(* IEC 61131-3 sources: daoli-st-library/DL_MathData (part 2) *)

(* ---- FC_DL_DtlStringConv.st ---- *)
(*
  ==================================================================
  组件名 Component  : FC_DL_DtlStringConv
  分类   Category   : DL_MathData
  复杂度 Complexity  : 中
  版本   Version    : 1.0.0
  功能   Purpose    : 日期时间 ↔ ASCII 串双向转换。定长 19 字符格式
                      'YYYY-MM-DD HH:MM:SS'。eStrToComp：串 → 六分量（分隔符
                      与数字位逐一校验，FIND 数字表解码）；eCompToStr：六分量
                      → 串（数字查表装配）。超长按 19 截断评估并置 bTrunc
                      （255 截断标志语义：入串超库上限 255 或超定长均置位）。
                      LGF Converter 组 DTL↔String 语义 clean-room。
  来源   Source     : T2-1-lgf-converter（LGF Converter 组 DTL↔String 语义）
  溯源   Origin     : 定长日期串装配/解析为公开工程语义，clean-room 自研实现，
                      未复制 LGF 或任何厂商私有库源码。
  平台   Platform   : 纯 IEC 61131-3（Standard.library: LEN / MID / CONCAT /
                      FIND，无私有库）
  分工声明 Split     : 与 FC_DL_AsciiFrameParse 分工——后者做 STX/ETX 仪表
                      帧解析，本件做定长日期时间串双向转换。
  作者   Author     : 道莅代码库 · PLC 编程专家（R59）
  ------------------------------------------------------------------
  边界 Boundary     :
                      一 值域闸（eCompToStr）：年 1970..2999 / 月 1..12 /
                         日 1..31 / 时 0..23 / 分秒 0..59，越域置 bError；
                      二 格式闸（eStrToComp）：定长 19、分隔符位置（5/8 =
                         '-'，11 = ' '，14/17 = ':'）、数字位非数字 → bError；
                      三 255 截断标志：LEN > 19 按前 19 位截断评估并置
                         bTrunc（信息级），LEN > 255 直接置 bError；
                      四 无除法无浮点（纯整数与串操作，无除零/非有限风险）；
                      五 无全局变量、无外部变量声明、无物理地址寻址。
  修订记录 Revision  :
    2026-11-21  v1.0.0  R59 首版（批 2 · 序号 6）
  ==================================================================
*)

TYPE E_DL_DtcMode :
(
    eStrToComp := 0, // 串 → 六分量 / the string to components direction
    eCompToStr := 1  // 六分量 → 串 / the components to string direction
);
END_TYPE

FUNCTION FC_DL_DtlStringConv : BOOL
VAR_INPUT
    eMode   : E_DL_DtcMode; // 转换方向枚举 [-] / the conversion direction enum
    sIn     : STRING(255) := ''; // 入串（eStrToComp 方向）[-] / the input string, the to components entry
    nYear   : DINT := 2000; // 年分量 [年]，域 1970..2999，eCompToStr 方向 / the year component
    nMonth  : DINT := 1;    // 月分量 [月]，域 1..12 / the month component
    nDay    : DINT := 1;    // 日分量 [日]，域 1..31 / the day component
    nHour   : DINT := 0;    // 时分量 [时]，域 0..23 / the hour component
    nMinute : DINT := 0;    // 分分量 [分]，域 0..59 / the minute component
    nSecond : DINT := 0;    // 秒分量 [秒]，域 0..59 / the second component
END_VAR
VAR_OUTPUT
    sOut    : STRING(23) := ''; // 出串 'YYYY-MM-DD HH:MM:SS' [-] / the output string, the fixed format
    oYear   : DINT := 0;   // 年分量输出 [年] / the year outlet
    oMonth  : DINT := 0;   // 月分量输出 [月] / the month outlet
    oDay    : DINT := 0;   // 日分量输出 [日] / the day outlet
    oHour   : DINT := 0;   // 时分量输出 [时] / the hour outlet
    oMinute : DINT := 0;   // 分分量输出 [分] / the minute outlet
    oSecond : DINT := 0;   // 秒分量输出 [秒] / the second outlet
    bValid  : BOOL := FALSE; // 结果可用标志 [-] / the result usable flag
    bTrunc  : BOOL := FALSE; // 截断标志（入串超定长 19 按前 19 位评估）[-] / the truncation flag, the long input evaluated by the first nineteen
    bError  : BOOL := FALSE; // 故障标志（格式/值域/超 255）[-] / the fault flag
END_VAR
VAR CONSTANT
    DL_DTC_DIGITS : STRING(10) := '0123456789'; // 数字字符表（FIND 解码基准）/ the digit table for the FIND decoding
    DL_DTC_LENFIX : DINT := 19; // 定长 [字符] / the fixed length
    DL_DTC_LENMAX : DINT := 255; // 库串上限 [字符] / the library string cap
END_VAR
VAR
    nLen   : DINT;  // 入串长度 [字符] / the input length
    sCh    : STRING(1); // 单字符工作量 [-] / the one char work value
    nPos   : DINT;  // 字表命中位（0 = 非数字）[位] / the table hit position, zero means non digit
    nI     : DINT;  // 数字位遍历索引 [位] / the digit position index
    nJ     : DINT;  // 字段遍历索引 [个] / the field index
    nVal   : DINT;  // 字段解析值工作量 [-] / the field parsed value work
    nDiv   : DINT;  // 位除子工作量（10 的幂，DINT 整除取位）[-] / the digit divisor, a power of ten
    aVal   : ARRAY[0..5] OF DINT; // 六分量装配工作数组 / the six component work array
    aField : ARRAY[0..5] OF DINT; // 六字段起始位组（1 基）/ the six field start positions, one based
    aWidth : ARRAY[0..5] OF DINT; // 六字段宽度组 [字符] / the six field widths
    aSep   : ARRAY[0..5] OF STRING(1); // 字段间分隔符组（末项空）/ the separators, the last empty
    bNeg   : BOOL;  // 保留（本件无符号语义，恒假）[-] / reserved, constant false
END_VAR

// 段 1｜返回值与输出预置（四段式第一段，R45）/ segment 1, preset the return and the outputs
FC_DL_DtlStringConv := FALSE; // 受理预置假 / preset the accepted false
sOut := ''; // 出串预置空 / preset the output empty
oYear := 0; oMonth := 0; oDay := 0; // 分量输出预置零 / preset the outlets zero
oHour := 0; oMinute := 0; oSecond := 0; // 分量输出预置零 / preset the outlets zero
bValid := FALSE; // 有效预置假 / preset the valid false
bTrunc := FALSE; // 截断预置假 / preset the trunc false
bError := FALSE; // 故障预置假 / preset the fault false
bNeg := FALSE; // 保留位恒假 / the reserved constant false

// 段 2｜方向一：串 → 六分量（格式闸 + 数字表解码 + 值域闸）/ segment 2, the string to components direction
IF eMode = E_DL_DtcMode.eStrToComp THEN // 方向一受理 / the direction one
    nLen := LEN(sIn); // 取长 / take the length
    IF nLen > DL_DTC_LENMAX THEN // 超 255 库上限：故障级 / beyond the cap, fault grade
        bError := TRUE; // 置故障 / raise the fault
        RETURN; // 早退 / return early
    END_IF
    IF nLen > DL_DTC_LENFIX THEN // 超定长：按前 19 位截断评估（信息级）/ beyond the fixed length, evaluate by the head
        bTrunc := TRUE; // 置截断标志 / raise the truncation
    ELSIF nLen < DL_DTC_LENFIX THEN // 短于定长：格式故障 / shorter than the fixed length
        bError := TRUE; // 置故障 / raise the fault
        RETURN; // 早退 / return early
    END_IF
    aField[0] := 1;  aWidth[0] := 4; // 年字段 YYYY / the year field
    aField[1] := 6;  aWidth[1] := 2; // 月字段 MM / the month field
    aField[2] := 9;  aWidth[2] := 2; // 日字段 DD / the day field
    aField[3] := 12; aWidth[3] := 2; // 时字段 HH / the hour field
    aField[4] := 15; aWidth[4] := 2; // 分字段 MI / the minute field
    aField[5] := 18; aWidth[5] := 2; // 秒字段 SS / the second field
    FOR nJ := 0 TO 5 DO // 逐字段解析 / per field parse
        nVal := 0; // 字段值清零 / clear the field value
        FOR nI := 0 TO aWidth[nJ] - 1 DO // 逐数字位 / per digit position
            sCh := MID(sIn, 1, aField[nJ] + nI); // 取单字符 / take one char
            nPos := FIND(DL_DTC_DIGITS, sCh); // 字表命中位 / the table hit position
            IF nPos = 0 THEN // 非数字字符 / a non digit char
                bError := TRUE; // 置故障（非法字符闸）/ raise the fault
                RETURN; // 早退 / return early
            END_IF
            nVal := (nVal * 10) + (nPos - 1); // 十进制装配 / assemble the decimal
        END_FOR
        aVal[nJ] := nVal; // 记字段值 / store the field value
    END_FOR
    IF (MID(sIn, 1, 5) <> '-') OR (MID(sIn, 1, 8) <> '-')
    OR (MID(sIn, 1, 11) <> ' ') OR (MID(sIn, 1, 14) <> ':')
    OR (MID(sIn, 1, 17) <> ':') THEN // 分隔符位置闸 / the separator gates
        bError := TRUE; // 置故障 / raise the fault
        RETURN; // 早退 / return early
    END_IF
    IF (aVal[0] < 1970) OR (aVal[0] > 2999) OR (aVal[1] < 1) OR (aVal[1] > 12)
    OR (aVal[2] < 1) OR (aVal[2] > 31) OR (aVal[3] > 23)
    OR (aVal[4] > 59) OR (aVal[5] > 59) THEN // 值域闸（边界一）/ the value domain gates
        bError := TRUE; // 置故障 / raise the fault
        RETURN; // 早退 / return early
    END_IF
    oYear := aVal[0]; oMonth := aVal[1]; oDay := aVal[2]; // 分量出口 / the outlets
    oHour := aVal[3]; oMinute := aVal[4]; oSecond := aVal[5]; // 分量出口 / the outlets
    bValid := TRUE; // 结果可用 / the result usable
    FC_DL_DtlStringConv := TRUE; // 受理 / accept

// 段 3｜方向二：六分量 → 串（值域闸 + 数字查表装配）/ segment 3, the components to string direction
ELSIF eMode = E_DL_DtcMode.eCompToStr THEN // 方向二受理 / the direction two
    IF (nYear < 1970) OR (nYear > 2999) OR (nMonth < 1) OR (nMonth > 12)
    OR (nDay < 1) OR (nDay > 31) OR (nHour > 23) OR (nHour < 0)
    OR (nMinute > 59) OR (nMinute < 0) OR (nSecond > 59) OR (nSecond < 0) THEN // 值域闸（边界一）/ the value domain gates
        bError := TRUE; // 置故障 / raise the fault
        RETURN; // 早退 / return early
    END_IF
    aVal[0] := nYear; aVal[1] := nMonth; aVal[2] := nDay; // 装配值组 / load the values
    aVal[3] := nHour; aVal[4] := nMinute; aVal[5] := nSecond; // 装配值组 / load the values
    aField[0] := 4; aField[1] := 2; aField[2] := 2; // 宽度组 / the widths
    aField[3] := 2; aField[4] := 2; aField[5] := 2; // 宽度组 / the widths
    aSep[0] := '-'; aSep[1] := '-'; aSep[2] := ' '; // 分隔符组 / the separators
    aSep[3] := ':'; aSep[4] := ':'; aSep[5] := '';  // 分隔符组（末项空）/ the separators, the last empty
    sOut := ''; // 出串清零 / clear the output
    FOR nJ := 0 TO 5 DO // 逐字段装配 / per field assembly
        sOut := CONCAT(sOut, aSep[nJ]); // 先接分隔符 / append the separator first
        nDiv := 1; // 位除子起步（10^(宽-1)）/ the divisor starts at one
        FOR nI := 1 TO aField[nJ] - 1 DO // 宽度减一次乘十 / the width minus one multiplies by ten
            nDiv := nDiv * 10; // 除子推进 / advance the divisor
        END_FOR
        FOR nI := 1 TO aField[nJ] DO // 高位到低位逐位 / per digit from the high position down
            sCh := MID(DL_DTC_DIGITS, 1, ((aVal[nJ] / nDiv) MOD 10) + 1); // DINT 整除取位查表（无浮点无 EXPT）/ the DINT divide and pick by the table
            sOut := CONCAT(sOut, sCh); // 接字符 / append the char
            nDiv := nDiv / 10; // 除子降位 / drop the divisor one decade
        END_FOR
    END_FOR
    bValid := TRUE; // 结果可用 / the result usable
    FC_DL_DtlStringConv := TRUE; // 受理 / accept
ELSE // 非法方向枚举兜底 / the illegal direction fallback
    bError := TRUE; // 置故障 / raise the fault
END_IF
END_FUNCTION

(* ---- FC_DL_DynViscosityUnitConvert.st ---- *)
(*==============================================================================
 * 组件名称 (Component)  : FC_DL_DynViscosityUnitConvert
 * 所属子库 (Sublibrary) : DL_MathData ｜ 版本 (Version) : 1.0.0 ｜ 2026-11-23
 * 兼容性   (Platform)   : CODESYS 3.5+ / TwinCAT 3 / 汇川 InoProShop / 施耐德 Machine Expert
 *                         仅依赖 IEC 61131-3 算术运算符，零厂商私有库
 * 功能描述 (Function)   : 动力粘度（dynamic viscosity，绝对粘度）单位互转，系数表驱动：
 *                         以 Pa·s 为中介单位，fHub = fValue × kSrc，fResult = fHub ÷ kDst；
 *                         系数为编译期非零常量，纯常量除法，结构性无除零。
 *                         **单位恒等说明**：1 cP ≡ 1 mPa·s（厘泊定义即毫帕·秒，两者为同一
 *                         物理量的两种书写），故两成员系数均为 1.0E-3；保留两个枚举成员
 *                         仅为适配不同 HMI 标签与协议字段，避免上游做字符串映射。
 *                         **与运动粘度的分工（关键）**：动力粘度 [Pa·s] 与运动粘度 [m²/s]
 *                         差一个密度因子（ν = η / ρ），本件不做该换算；运动粘度件为
 *                         FC_DL_ViscosityUnitConvert（mm²/s 族）。
 *                         负粘度物理上不存在 → 故障级 eNegativeValue 拒绝（不取绝对值）。
 * 接口     (Interface)  : 输入 fValue 被换算动力粘度 [源单位]、eSrc 源单位、eDst 目标单位；
 *                         输出 fConverted 换算结果 [目标单位]、eErrCode（E_DL_DynViscConvErr）；
 *                         返回值 = 数值可信标志。
 * 边界     (Boundary)   : ① 单位枚举越域 → 故障级 eInvalidUnit，结果哨兵 0。
 *                         ② 非有限双判（NaN / ±Inf），命中即故障级 eNonFinite。
 *                         ③ 负粘度 → 故障级 eNegativeValue（拒绝换算）。
 *                         ④ 零粘度 → 信息级 eZeroValue（物理上仅真空 / 静止，多为未充油），
 *                            结果仍可信并返回 TRUE（0 Pa·s = 0 cP 恒成立）。
 *                         ⑤ 中介值与结果各复检一次（四段式第四段）。
 *                         ⑥ 温度不补偿：动力粘度强依赖温度，本件为纯量纲换算，
 *                            调用方必须保证参与比较的数据同温基准（推荐 40 ℃）。
 *                         ⑦ 零全局耦合（无 GVL / VAR_EXTERNAL / 物理地址）。
 * 码表     (Codes)      : 本件不占用全局数字码位（R297 零码位范式）；出口为 BOOL + LREAL +
 *                         本文件内 enum E_DL_DynViscConvErr（全库唯一属主）。
 * 分工声明 (Scope)      : 运动粘度归 FC_DL_ViscosityUnitConvert（E_DL_ViscUnit 属主）；
 *                         粘度-温度曲线拟合与油品换油判定不在本件范围。
 * 归属     (Ownership)  : E_DL_DynViscUnit / E_DL_DynViscConvErr 归属本文件（全库唯一属主，R264）。
 * 红线自检 (Redline)    : R1 ✓ 零 GVL ｜ R2 ✓ 零 %I/%Q ｜ R3 ✓ 纯 IEC ｜ R4 ✓ 非有限双判 +
 *                         CASE ELSE 兜底 + 常量除法无除零 + 负值闸 ｜ R5 ✓ 逐行同行双语注释
 *                         R6 ✓ CASE ELSE 兜底 ｜ R7 N/A（无实例调用）
 * 修订历史 (Revision)   : 2026-11-23  v1.0.0  R78-B2 首版（因 FC_DL_ViscosityUnitConvert
 *                         名称为运动粘度件占用，本件按动力粘度口径另立名）
 * 验收向量 (Acceptance) :
 *   A1 fValue=1000.0, eSrc=eCp, eDst=ePas → 1.0（容差 1E-12）；
 *   A2 fValue=1.0, eSrc=ePas, eDst=eCp → 1000.0；
 *   A3 fValue=1.0, eSrc=eCp, eDst=eMPas → 1.0（恒等关系）；
 *   A4 fValue=-5.0, eSrc=eCp, eDst=ePas → 0 哨兵, eNegativeValue, 返回 FALSE；
 *   A5 fValue=0.0, eSrc=ePas, eDst=eCp → 0.0, eZeroValue, 返回 TRUE。
 *============================================================================*)

(*-----------------------------------------------------------------------------
 * 枚举: E_DL_DynViscUnit（动力粘度单位表，归属本文件，全库唯一属主）
 *----------------------------------------------------------------------------*)
TYPE E_DL_DynViscUnit :
(
    ePas  := 0,   // 帕斯卡秒（中介单位，SI 一致单位） / Pascal second, hub unit
    eCp   := 1,   // 厘泊（= 1.0E-3 Pa·s） / Centipoise, equals 1.0E-3 Pa s
    eMPas := 2    // 毫帕秒（= 1.0E-3 Pa·s，与厘泊恒等） / Millipascal second, identical to centipoise
);
END_TYPE

(*-----------------------------------------------------------------------------
 * 枚举: E_DL_DynViscConvErr（动力粘度换算出口码；信息级 = 0..9，故障级 = 10 起）
 *----------------------------------------------------------------------------*)
TYPE E_DL_DynViscConvErr :
(
    eOk            := 0,   // 信息级：换算完成 / Info: conversion completed
    eZeroValue     := 1,   // 信息级：零粘度（多为未充油） / Info: zero viscosity, result still trustworthy
    eInvalidUnit   := 10,  // 故障级：单位枚举越域 / Fault: unit enum out of domain
    eNonFinite     := 11,  // 故障级：输入或结果非有限 / Fault: non-finite input or result
    eNegativeValue := 12   // 故障级：负粘度 / Fault: negative viscosity
);
END_TYPE

FUNCTION FC_DL_DynViscosityUnitConvert : BOOL
VAR_INPUT
    fValue : LREAL;             // 被换算动力粘度 [源单位] / Dynamic viscosity value in the source unit
    eSrc   : E_DL_DynViscUnit;  // 源单位枚举 [-] / Source unit enum
    eDst   : E_DL_DynViscUnit;  // 目标单位枚举 [-] / Destination unit enum
END_VAR
VAR_OUTPUT
    fConverted : LREAL;                 // 换算结果 [目标单位] / Converted result in the destination unit
    eErrCode   : E_DL_DynViscConvErr;   // 出口码 [-] / Outlet code
END_VAR
VAR
    _bBadValue : BOOL;   // 输入非有限标志 [-] / Non-finite input flag
    _fHub      : LREAL;  // 中介动力粘度 [Pa·s] / Hub dynamic viscosity in pascal second
END_VAR
VAR CONSTANT
    DL_DVC_ZERO : LREAL := 0.0;       // 零基准与零值判定基准 [-] / Zero base
    DL_DVC_PAS  : LREAL := 1.0;       // Pa·s → Pa·s 恒等系数 [-] / Hub identity factor
    DL_DVC_CP   : LREAL := 1.0E-3;    // cP → Pa·s 换算系数 [-] / Centipoise factor
    DL_DVC_MPAS : LREAL := 1.0E-3;    // mPa·s → Pa·s 换算系数 [-] / Millipascal second factor
    DL_DVC_EPS  : LREAL := 1.0E-12;   // 零值判定容差 [-] / Zero-detection tolerance
END_VAR

(* —— 段 0：出口预置安全侧 —— *)
FC_DL_DynViscosityUnitConvert := FALSE;              // 返回值预置不可信 / Return preset not trustworthy
fConverted := DL_DVC_ZERO;                           // 结果哨兵 0 / Result sentinel
eErrCode   := E_DL_DynViscConvErr.eInvalidUnit;      // 预置最严码 / Preset strictest code

(* —— 段 1：非有限域闸（R79 双判） —— *)
_bBadValue := (fValue <> fValue) OR ((fValue - fValue) <> DL_DVC_ZERO);      // 输入非有限 / Input non-finite
IF _bBadValue THEN
    eErrCode := E_DL_DynViscConvErr.eNonFinite;      // 故障级码 / Fault-level code
    RETURN;
END_IF

(* —— 段 2：负粘度域闸（零值放行，由段 6 置信息码） —— *)
IF fValue < DL_DVC_ZERO THEN
    eErrCode := E_DL_DynViscConvErr.eNegativeValue;  // 故障级码 / Fault-level code
    RETURN;
END_IF

(* —— 段 3：源单位 → 中介 Pa·s（CASE ELSE 拦截越域） —— *)
CASE eSrc OF
    E_DL_DynViscUnit.ePas :
        _fHub := fValue * DL_DVC_PAS;                // 直通 / Hub pass-through
    E_DL_DynViscUnit.eCp :
        _fHub := fValue * DL_DVC_CP;                 // cP × 1E-3 / Centipoise scaled
    E_DL_DynViscUnit.eMPas :
        _fHub := fValue * DL_DVC_MPAS;               // mPa·s × 1E-3 / Millipascal second scaled
ELSE
    _fHub    := DL_DVC_ZERO;                         // 中介值回哨兵 / Hub back to sentinel
    eErrCode := E_DL_DynViscConvErr.eInvalidUnit;    // 故障级：源单位越域 / Fault: source out of domain
    RETURN;
END_CASE

(* —— 段 4：中介 Pa·s → 目标单位（除数为常量，均非零） —— *)
CASE eDst OF
    E_DL_DynViscUnit.ePas :
        fConverted := _fHub / DL_DVC_PAS;            // ÷1 / Divide by identity
    E_DL_DynViscUnit.eCp :
        fConverted := _fHub / DL_DVC_CP;             // ÷1E-3 / Divide by centipoise factor
    E_DL_DynViscUnit.eMPas :
        fConverted := _fHub / DL_DVC_MPAS;           // ÷1E-3 / Divide by millipascal second factor
ELSE
    fConverted := DL_DVC_ZERO;                       // 结果回哨兵 / Result back to sentinel
    eErrCode   := E_DL_DynViscConvErr.eInvalidUnit;  // 故障级：目标单位越域 / Fault: destination out of domain
    RETURN;
END_CASE

(* —— 段 5：中介值与结果复检（四段式第四段） —— *)
IF (_fHub <> _fHub) OR ((_fHub - _fHub) <> DL_DVC_ZERO)
    OR (fConverted <> fConverted) OR ((fConverted - fConverted) <> DL_DVC_ZERO) THEN
    fConverted := DL_DVC_ZERO;                       // 复检异常回哨兵 / Recheck failed: sentinel
    eErrCode   := E_DL_DynViscConvErr.eNonFinite;    // 故障级码 / Fault-level code
    RETURN;
END_IF

(* —— 段 6：成功出口（零值单列信息码，提示上游可能未充油） —— *)
IF (fValue < DL_DVC_EPS) AND (fValue > -DL_DVC_EPS) THEN
    eErrCode := E_DL_DynViscConvErr.eZeroValue;      // 信息级：零粘度 / Info: zero viscosity
ELSE
    eErrCode := E_DL_DynViscConvErr.eOk;             // 信息级：换算完成 / Info: conversion completed
END_IF
FC_DL_DynViscosityUnitConvert := TRUE;               // 换算有效 / Conversion valid
END_FUNCTION

(* ---- FC_DL_EnergyUnitConvert.st ---- *)
(*==============================================================================
 * 组件名称 (Component)  : FC_DL_EnergyUnitConvert
 * 所属子库 (Sublibrary) : DL_MathData
 * 当前版本 (Version)    : 1.0.0
 * 兼容性   (Platform)   : CODESYS 3.5+ / TwinCAT 3 / 汇川 InoProShop / 施耐德 Machine Expert
 *                         仅依赖 IEC 61131-3 算术运算符，零厂商私有库
 * 功能描述 (Function)   : 能量单位换算（系数表驱动）：以千焦（kJ）为中介单位，
 *                         fHub = fValue × kSrc，fResult = fHub ÷ kDst；系数为编译期
 *                         非零常量，纯常量除法，结构性无除零。
 *                         **符号语义**：能量允许负值（电能回馈 / 热流反向 / 净能耗为负），
 *                         故本件**不做负值拒绝**，仅在结果非有限时兜底。此点与
 *                         长度/质量/体积等几何量件不同，属显式量纲差异，已在此声明。
 *                         口径：cal 取热化学卡（4.1868 J）；BTU 取 IT 表（1055.05585262 J）。
 * 接口     (Interface)  : 输入 fValue 被换算能量 [源单位]、eSrc 源单位、eDst 目标单位；
 *                         输出 fConverted 换算结果 [目标单位]、eErrCode（E_DL_EnergyConvErr）；
 *                         返回值 = bValid 数值可信标志（TRUE = fConverted 可信）。
 * 边界     (Boundary)   : ① 属主边界：只做单位换算，不做累计电量计费、不做峰谷分段统计。
 *                         ② 单位枚举越域 → 故障级 eInvalidUnit，结果哨兵 0。
 *                         ③ 非有限双判，命中即故障级 eNonFinite。
 *                         ④ 负值合法（回馈 / 反向），不置任何码。
 *                         ⑤ 零值 → 信息级 eZeroValue。
 *                         ⑥ kJ ↔ kWh 跨越 3600 倍，结果复检防非有限。
 *                         ⑦ 零全局耦合（无 GVL / VAR_EXTERNAL / 物理地址）。
 * 分工声明 (Scope)      : 与 `FC_DL_PowerUnitConvert` 分工：功率是能量对时间的导数，
 *                         能量累计与功率积分（含时基）归调用方的累计 FB，本件不内联时间。
 * 来源标签 (Source Tag) : 开源溯源：lgf-math 换算系数（公开物理常数，clean-room 重写）；许可证 MIT（仅参考语义，代码原创）
 * 码表     (Codes)      : 本件不占用全局数字码位；出口为 BOOL + LREAL +
 *                         本文件内定义 enum E_DL_EnergyConvErr（全库唯一）。
 * 红线自检 (Redline)    : R1 ✓ 零 GVL/VAR_EXTERNAL ｜ R2 ✓ 零 %I/%Q/%M ｜ R3 ✓ 纯 IEC 61131-3
 *                         R4 ✓ 非有限双判 + 枚举域闸 + 常量除法无除零（负值按量纲放行） ｜ R5 ✓ 声明逐行同行双语注释
 *                         R6 N/A（纯函数无状态机） ｜ R7 N/A（无实例调用）
 * 修订历史 (Revision)   : 2026-11-23  v1.0.0  R77 首版（批次 B2 · 序号 17）
 * 验收向量 (Acceptance) : ① fValue=1.0, eSrc=eKwh, eDst=eKj → 1×3600 = 3600.0 kJ, eOk, TRUE；
 *                         ② fValue=4186.8, eSrc=eKj, eDst=eCal → 4186.8×1.0 = 4186.8 kJ,
 *                         ÷0.0041868 = 1000000.0 cal（容差 1E-3）；
 *                         ③ fValue=1.0, eSrc=eBtu, eDst=eKj → 1.05505585262 kJ（容差 1E-12）；
 *                         ④ fValue=-2.5, eSrc=eKwh, eDst=eKj → -9000.0 kJ（负值合法）, eOk, TRUE；
 *                         ⑤ fValue=0.0, eSrc=eKj, eDst=eKwh → 0.0, 返回 TRUE, eZeroValue。
 *==============================================================================*)

(*-----------------------------------------------------------------------------
 * 枚举: E_DL_EnergyUnit（能量单位表，归属 DL_MathData，与本件同文件，全库唯一属主）
 *----------------------------------------------------------------------------*)
TYPE E_DL_EnergyUnit :
(
    eKj   := 0,   // 千焦（中介单位） / Kilojoule, hub unit
    eKwh  := 1,   // 千瓦时（= 3600 kJ） / Kilowatt hour
    eCal  := 2,   // 卡（热化学卡，= 0.0041868 kJ） / Thermochemical calorie
    eBtu  := 3    // 英热单位（IT 表，= 1.05505585262 kJ） / British thermal unit, IT table
);
END_TYPE

(*-----------------------------------------------------------------------------
 * 枚举: E_DL_EnergyConvErr（能量换算错误码）
 * 分级: 本件无「负值」故障码——能量负值属合法物理语义（回馈/反向）。
 *----------------------------------------------------------------------------*)
TYPE E_DL_EnergyConvErr :
(
    eOk        := 0,   // 信息级：换算完成 / Info: conversion completed
    eZeroValue := 1,   // 信息级：输入为零（合法） / Info: zero input, legal
    eInvalidUnit := 2, // 故障级：单位枚举越域 / Fault: unit enum out of domain
    eNonFinite := 3    // 故障级：输入非有限 / Fault: non-finite input
);
END_TYPE

FUNCTION FC_DL_EnergyUnitConvert : BOOL
VAR_INPUT
    fValue : LREAL;            // 被换算能量值（可负） [源单位] / Energy value, negative allowed, in source unit
    eSrc   : E_DL_EnergyUnit;  // 源单位枚举 [-] / Source unit enum
    eDst   : E_DL_EnergyUnit;  // 目标单位枚举 [-] / Destination unit enum
END_VAR
VAR_OUTPUT
    fConverted : LREAL;              // 换算结果（可负） [目标单位] / Converted result, may be negative
    eErrCode   : E_DL_EnergyConvErr; // 错误码出口 [-] / Error code outlet
END_VAR
VAR
    _bNonFin : BOOL;   // 输入非有限当拍标志 [-] / Non-finite input flag
    _fHub    : LREAL;  // 中介能量值 [kJ] / Hub energy value in kilojoules
END_VAR
VAR CONSTANT
    DL_EUC_KJ   : LREAL := 1.0;             // kJ → kJ 恒等系数 [-] / Hub identity factor
    DL_EUC_KWH  : LREAL := 3600.0;          // kWh → kJ 换算系数 [kJ/kWh] / Kilowatt hour to kilojoule factor
    DL_EUC_CAL  : LREAL := 0.0041868;       // cal → kJ 换算系数 [kJ/cal] / Calorie to kilojoule factor
    DL_EUC_BTU  : LREAL := 1.05505585262;   // BTU(IT) → kJ 换算系数 [kJ/BTU] / BTU to kilojoule factor
    DL_EUC_ZERO : LREAL := 0.0;             // 零值与非有限判零基准 [-] / Zero and non-finite base
END_VAR

(* —— 段 0：出口预置安全值 —— *)
FC_DL_EnergyUnitConvert := FALSE;                  // 返回值预置无效 / Return preset invalid
fConverted := DL_EUC_ZERO;                         // 结果哨兵 0 / Result sentinel
eErrCode   := E_DL_EnergyConvErr.eInvalidUnit;     // 预置最严码 / Preset strictest code

(* —— 段 1：非有限域闸（R79 双判） —— *)
_bNonFin := (fValue <> fValue) OR ((fValue - fValue) <> DL_EUC_ZERO);   // 非有限判定 / Non-finite test
IF _bNonFin THEN
    eErrCode := E_DL_EnergyConvErr.eNonFinite;     // 故障级码 / Fault-level code
    RETURN;
END_IF

(* —— 段 2：极性说明（能量负值合法，本段仅注释占位，不做拦截） —— *)
(* Negative energy is physically legal, so no polarity gate is applied here. *)

(* —— 段 3：源单位 → 中介 kJ —— *)
IF eSrc = E_DL_EnergyUnit.eKj THEN
    _fHub := fValue * DL_EUC_KJ;                   // 直通 / Hub pass-through
ELSIF eSrc = E_DL_EnergyUnit.eKwh THEN
    _fHub := fValue * DL_EUC_KWH;                  // kWh × 3600 / Kilowatt hour scaled
ELSIF eSrc = E_DL_EnergyUnit.eCal THEN
    _fHub := fValue * DL_EUC_CAL;                  // cal × 0.0041868 / Calorie scaled
ELSIF eSrc = E_DL_EnergyUnit.eBtu THEN
    _fHub := fValue * DL_EUC_BTU;                  // BTU × 1.05505585262 / BTU scaled
ELSE
    RETURN;                                        // 源单位越域 / Source unit out of domain
END_IF

(* —— 段 4：中介 kJ → 目标单位（常量除法，分母非零） —— *)
IF eDst = E_DL_EnergyUnit.eKj THEN
    fConverted := _fHub / DL_EUC_KJ;               // ÷1 / Divide by identity
ELSIF eDst = E_DL_EnergyUnit.eKwh THEN
    fConverted := _fHub / DL_EUC_KWH;              // ÷3600 / Divide by kilowatt hour factor
ELSIF eDst = E_DL_EnergyUnit.eCal THEN
    fConverted := _fHub / DL_EUC_CAL;              // ÷0.0041868 / Divide by calorie factor
ELSIF eDst = E_DL_EnergyUnit.eBtu THEN
    fConverted := _fHub / DL_EUC_BTU;              // ÷1.05505585262 / Divide by BTU factor
ELSE
    eErrCode   := E_DL_EnergyConvErr.eInvalidUnit; // 目标单位越域 / Destination out of domain
    fConverted := DL_EUC_ZERO;
    RETURN;
END_IF

(* —— 段 5：结果非有限复检兜底 —— *)
IF (fConverted <> fConverted) OR ((fConverted - fConverted) <> DL_EUC_ZERO) THEN
    fConverted := DL_EUC_ZERO;                     // 复检异常回哨兵 / Recheck failed: sentinel
    eErrCode   := E_DL_EnergyConvErr.eNonFinite;   // 故障级码 / Fault-level code
    RETURN;
END_IF

(* —— 段 6：成功出口 —— *)
IF fValue = DL_EUC_ZERO THEN
    eErrCode := E_DL_EnergyConvErr.eZeroValue;     // 信息级：零值 / Info: zero value
ELSE
    eErrCode := E_DL_EnergyConvErr.eOk;            // 信息级成功 / Info success
END_IF
FC_DL_EnergyUnitConvert := TRUE;                   // 换算有效 / Conversion valid

END_FUNCTION

(* ---- FC_DL_FiniteClassify.st ---- *)
(*
    FC_DL_FiniteClassify —— LREAL 非有限分类原子
    ------------------------------------------------------------------
    组件名称  : FC_DL_FiniteClassify
    分类      : DL_MathData / FloatFiniteness
    前缀      : FC_DL_
    版本      : 1.0.0
    溯源      : IEC 61131-3 标准语义的道莅防御性实现（IEEE 754 NaN 自反性
                与 Inf 差值自反判据的原子化提取，判据即库内 R79 非有限
                双判的语义本体）；实现 / 引脚名 / 枚举 100% 自有；
                clean-room 声明 —— 零代码行复制，无闭源参考。
    平台      : 纯 IEC 61131-3（LREAL 比较 + 标准 ABS），无内建函数依赖，
                CODESYS 3.5 / TwinCAT 3 / InoProShop / Machine Expert 通用
    作者      : 道莅代码库 · PLC编程专家（R72 构建轮 · 批 1 · 序号 2）
    ------------------------------------------------------------------
    功能说明  : 把散落在库内各件的内联 R79 非有限判据提取为**全库首个
                非有限分类属主**，输出 IEEE 754 语义四态：eFinite / ePosInf /
                eNegInf / eNaN，并给 bFinite 布尔快照。真实工况：闸前置
                分类诊断文本（HMI 显示「断线 / 无穷 / 正常」）、诊断日志分桶。
                判据链（禁近似阈值，R79）：
                ① NaN 用自反性 x <> x 判（NaN 与任何值比较均为 FALSE，含自身）；
                ② Inf 用差值自反判 (x − x) <> 0（有限值差恒为 0，无穷处产 NaN），
                   判出后按符号二分（x > 0.0 → ePosInf，x < 0.0 → eNegInf；
                   x = 0.0 在非 NaN 前提下差值必为 0，不会落入本分支）；
                ③ 其余 eFinite。
                幅值常量 1.7976931348623157E308 只可作注释旁证（LREAL 最大
                有限值），**不得作为判据**——近似阈值会在 [近似值, 真实最大值]
                区间制造假阳性带（R79 教训）。
                与库内各件内联 R79 判据的关系 = 「原子提取」而非语义变更：
                各件可组合调用本件但不强制回改存量（存量回改挂账不改码，
                R333 口径）。本件不做幅值上界筛查——上界筛查属调用方业务
                语义，本件只分 IEEE 语义四态。
    错误码    : N/A —— 本件为全定义域全值函数（任何 LREAL 入参都得到确定
                分类），无故障 / 信息出口，无码位分配。
    码位总账  : 无（全值函数，四态穷尽 LREAL 全域）
    状态机    : N/A —— 纯函数无状态，无 CASE 可写，非法状态不可能出现
    边界与披露: 一 无定时器 / 无沿检测实例 / 无数组下标 / 无除法 / 无循环，
                   零除零面与死循环面，周期安全规则 N/A；
                二 零全局变量、零 VAR_EXTERNAL、零物理地址；
                三 验收向量：V1 1.0 → eFinite + bFinite=TRUE；
                   V2 0.0 / 0.0（NaN）→ eNaN + bFinite=FALSE；
                   V3 1.0 / 0.0（+Inf）→ ePosInf + bFinite=FALSE；
                   V4 −1.0 / 0.0（−Inf）→ eNegInf + bFinite=FALSE；
                   V5 −0.0 → eFinite（负零是有限值，差值恒 0）。
                算法已证（脚本）：未跑 ｜ 编译器已证（三平台）：未跑
    修订记录  : 2026-11-23 v1.0.0 首次入库（R72 构建轮 · 批 1 · 序号 2）
*)
TYPE E_DL_FiniteKind :
(
    eFinite := 0,                          // 有限值：正常数值 / finite, a normal numeric value
    ePosInf := 1,                          // 正无穷：+Inf，多为除零 / 上溢 / the positive infinity
    eNegInf := 2,                          // 负无穷：−Inf，多为下溢 / 负向除零 / the negative infinity
    eNaN    := 3                           // 非数：断线 / 无效运算结果 / the not a number class
);
END_TYPE

FUNCTION FC_DL_FiniteClassify : E_DL_FiniteKind
VAR_INPUT
    fVal : LREAL;                          (* 待分类值，[任意物理量纲，无量纲语义]，本件不解释量纲 / the value under test, dimension free, the FC never interprets units *)
END_VAR
VAR_OUTPUT
    bFinite : BOOL;                        (* 有限值快照：TRUE 当且仅当分类为 eFinite / the finite snapshot, TRUE iff eFinite *)
END_VAR

// 段 1｜返回值与状态预置（统一出口预置，R256）/ segment 1, preset the return and the status
FC_DL_FiniteClassify := E_DL_FiniteKind.eFinite; // 预置有限分类 / preset the finite class
bFinite := FALSE;                        // 预置非有限快照（段 3 正常出口翻转）/ preset the snapshot false

// 段 2｜NaN 自反判（NaN 与自身比较为 FALSE，R79 判据一）/ segment 2, the NaN reflexive test
IF fVal <> fVal THEN                     // 自比较为假即 NaN / a false self comparison means NaN
    FC_DL_FiniteClassify := E_DL_FiniteKind.eNaN; // 分类非数 / classify NaN
    bFinite := FALSE;                    // 快照非有限 / the snapshot false
    RETURN;                              // 结构早退 / structural exit
END_IF

// 段 3｜Inf 差值自反判（有限值差恒 0，无穷处产 NaN，R79 判据二）+ 符号二分 / segment 3, the infinity difference test and the sign split
IF (fVal - fVal) <> 0.0 THEN             // 差值非零即无穷 / a non zero difference means infinity
    IF fVal > 0.0 THEN                   // 正无穷支（NaN 已在段 2 排除，0.0 不会落入本支）/ the positive branch
        FC_DL_FiniteClassify := E_DL_FiniteKind.ePosInf; // 分类正无穷 / classify plus infinity
    ELSE                                 // 负无穷支 / the negative branch
        FC_DL_FiniteClassify := E_DL_FiniteKind.eNegInf; // 分类负无穷 / classify minus infinity
    END_IF
    bFinite := FALSE;                    // 快照非有限 / the snapshot false
    RETURN;                              // 结构早退 / exit
END_IF

// 段 4｜有限值正常出口（旁证注释：LREAL 最大有限值 1.7976931348623157E308，
//        仅注释不作判据，R79 禁近似阈值）/ segment 4, the finite outlet
FC_DL_FiniteClassify := E_DL_FiniteKind.eFinite; // 分类有限 / classify finite
bFinite := TRUE;                         // 快照有限 / the snapshot true
END_FUNCTION

(* ---- FC_DL_FlowMassUnitConvert.st ---- *)
(*==============================================================================
 * 组件名称 (Component)  : FC_DL_FlowMassUnitConvert
 * 所属子库 (Sublibrary) : DL_MathData ｜ 版本 (Version) : 1.0.0 ｜ 2026-11-23
 * 兼容性   (Platform)   : CODESYS 3.5+ / TwinCAT 3 / 汇川 InoProShop / 施耐德 Machine Expert
 *                         仅依赖 IEC 61131-3 算术运算符，零厂商私有库
 * 功能描述 (Function)   : 质量流量单位互转（系数表驱动）：以 kg/h 为中介单位，
 *                         fHub = fValue × kSrc，fResult = fHub ÷ kDst；系数为编译期非零常量，
 *                         纯常量除法，结构性无除零。枚举源/目标越界由 CASE ... ELSE 拦截并
 *                         返回 0 哨兵。**与体积流量的分工**：本件只换质量流量，
 *                         体积流量（m³/h / L/min / SCFM）归 FC_DL_FlowUnitConvert；
 *                         两者之间的换算需介质密度，属组合换算，由调用方分两步完成。
 * 接口     (Interface)  : 输入 fValue 被换算质量流量 [源单位]、eSrc 源单位、eDst 目标单位；
 *                         输出 fConverted 换算结果 [目标单位]、eErrCode（E_DL_FlowMassConvErr）；
 *                         返回值 = 数值可信标志。
 * 边界     (Boundary)   : ① 质量流量可反向（倒罐 / 回流），负值合法，不设符号闸。
 *                         ② 单位枚举越域 → 故障级 eInvalidUnit，结果哨兵 0。
 *                         ③ 非有限双判，命中即故障级 eNonFinite。
 *                         ④ 中介值与结果各复检一次（四段式第四段）。
 *                         ⑤ 零值合法（停流），置信息级 eZeroValue。
 *                         ⑥ 换算系数为国际定义值：1 t = 1000 kg（公吨，非短吨）；
 *                            1 lb = 0.45359237 kg（国际磅，1959 约定值）。
 *                         ⑦ 零全局耦合（无 GVL / VAR_EXTERNAL / 物理地址）。
 * 码表     (Codes)      : 本件不占用全局数字码位（R297 零码位范式）；出口为 BOOL + LREAL +
 *                         本文件内 enum E_DL_FlowMassConvErr（全库唯一属主）。
 * 分工声明 (Scope)      : 体积流量归 FC_DL_FlowUnitConvert；质量/体积互转需密度，
 *                         本件不内联密度（R216 单一职责）。
 * 归属     (Ownership)  : E_DL_FlowMassUnit / E_DL_FlowMassConvErr 归属本文件（全库唯一属主，R264）。
 * 红线自检 (Redline)    : R1 ✓ 零 GVL ｜ R2 ✓ 零 %I/%Q ｜ R3 ✓ 纯 IEC ｜ R4 ✓ 非有限双判 +
 *                         CASE ELSE 兜底 + 常量除法无除零 ｜ R5 ✓ 逐行同行双语注释 ｜ R6 ✓ CASE ELSE
 *                         R7 N/A（无实例调用）
 * 修订历史 (Revision)   : 2026-11-23  v1.0.0  R78-B2 首版
 * 验收向量 (Acceptance) :
 *   A1 fValue=1.0, eSrc=eTH, eDst=eKgH → 1000.0；
 *   A2 fValue=1000.0, eSrc=eKgH, eDst=eTH → 1.0（容差 1E-12）；
 *   A3 fValue=1.0, eSrc=eLbH, eDst=eKgH → 0.45359237；
 *   A4 fValue=-250.0, eSrc=eKgH, eDst=eTH → -0.25（反向流合法）；
 *   A5 fValue=2.0, eSrc=非法值 9, eDst=eKgH → 0 哨兵, eInvalidUnit, 返回 FALSE。
 *============================================================================*)

(*-----------------------------------------------------------------------------
 * 枚举: E_DL_FlowMassUnit（质量流量单位表，归属本文件，全库唯一属主）
 *----------------------------------------------------------------------------*)
TYPE E_DL_FlowMassUnit :
(
    eKgH  := 0,   // 千克每小时（中介单位） / Kilogram per hour, hub unit
    eTH   := 1,   // 公吨每小时（= 1000 kg/h） / Metric tonne per hour, equals 1000 kg/h
    eLbH  := 2    // 磅每小时（= 0.45359237 kg/h） / Pound per hour, equals 0.45359237 kg/h
);
END_TYPE

(*-----------------------------------------------------------------------------
 * 枚举: E_DL_FlowMassConvErr（质量流量换算出口码；信息级 = 0..9，故障级 = 10 起）
 *----------------------------------------------------------------------------*)
TYPE E_DL_FlowMassConvErr :
(
    eOk          := 0,   // 信息级：换算完成 / Info: conversion completed
    eZeroValue   := 1,   // 信息级：零流量（停流） / Info: zero flow, result still trustworthy
    eInvalidUnit := 10,  // 故障级：单位枚举越域 / Fault: unit enum out of domain
    eNonFinite   := 11   // 故障级：输入或结果非有限 / Fault: non-finite input or result
);
END_TYPE

FUNCTION FC_DL_FlowMassUnitConvert : BOOL
VAR_INPUT
    fValue : LREAL;              // 被换算质量流量 [源单位] / Mass flow value in the source unit
    eSrc   : E_DL_FlowMassUnit;  // 源单位枚举 [-] / Source unit enum
    eDst   : E_DL_FlowMassUnit;  // 目标单位枚举 [-] / Destination unit enum
END_VAR
VAR_OUTPUT
    fConverted : LREAL;                 // 换算结果 [目标单位] / Converted result in the destination unit
    eErrCode   : E_DL_FlowMassConvErr;   // 出口码 [-] / Outlet code
END_VAR
VAR
    _bBadValue : BOOL;   // 输入非有限标志 [-] / Non-finite input flag
    _fHub      : LREAL;  // 中介质量流量 [kg/h] / Hub mass flow in kilogram per hour
END_VAR
VAR CONSTANT
    DL_FMC_ZERO : LREAL := 0.0;          // 零基准与零值判定基准 [-] / Zero base
    DL_FMC_KGH  : LREAL := 1.0;          // kg/h → kg/h 恒等系数 [-] / Hub identity factor
    DL_FMC_TH   : LREAL := 1000.0;       // t/h → kg/h 换算系数 [-] / Metric tonne per hour factor
    DL_FMC_LBH  : LREAL := 0.45359237;   // lb/h → kg/h 换算系数 [-] / Pound per hour factor
    DL_FMC_EPS  : LREAL := 1.0E-12;      // 零值判定容差 [-] / Zero-detection tolerance
END_VAR

(* —— 段 0：出口预置安全侧 —— *)
FC_DL_FlowMassUnitConvert := FALSE;                  // 返回值预置不可信 / Return preset not trustworthy
fConverted := DL_FMC_ZERO;                           // 结果哨兵 0 / Result sentinel
eErrCode   := E_DL_FlowMassConvErr.eInvalidUnit;     // 预置最严码 / Preset strictest code

(* —— 段 1：非有限域闸（R79 双判） —— *)
_bBadValue := (fValue <> fValue) OR ((fValue - fValue) <> DL_FMC_ZERO);      // 输入非有限 / Input non-finite
IF _bBadValue THEN
    eErrCode := E_DL_FlowMassConvErr.eNonFinite;     // 故障级码 / Fault-level code
    RETURN;
END_IF

(* —— 段 2：源单位 → 中介 kg/h（CASE ELSE 拦截越域） —— *)
CASE eSrc OF
    E_DL_FlowMassUnit.eKgH :
        _fHub := fValue * DL_FMC_KGH;                // 直通 / Hub pass-through
    E_DL_FlowMassUnit.eTH :
        _fHub := fValue * DL_FMC_TH;                 // t/h × 1000 / Metric tonne per hour scaled
    E_DL_FlowMassUnit.eLbH :
        _fHub := fValue * DL_FMC_LBH;                // lb/h × 0.45359237 / Pound per hour scaled
ELSE
    _fHub    := DL_FMC_ZERO;                         // 中介值回哨兵 / Hub back to sentinel
    eErrCode := E_DL_FlowMassConvErr.eInvalidUnit;   // 故障级：源单位越域 / Fault: source out of domain
    RETURN;
END_CASE

(* —— 段 3：中介 kg/h → 目标单位（除数为常量，均非零） —— *)
CASE eDst OF
    E_DL_FlowMassUnit.eKgH :
        fConverted := _fHub / DL_FMC_KGH;            // ÷1 / Divide by identity
    E_DL_FlowMassUnit.eTH :
        fConverted := _fHub / DL_FMC_TH;             // ÷1000 / Divide by metric tonne factor
    E_DL_FlowMassUnit.eLbH :
        fConverted := _fHub / DL_FMC_LBH;            // ÷0.45359237 / Divide by pound per hour factor
ELSE
    fConverted := DL_FMC_ZERO;                       // 结果回哨兵 / Result back to sentinel
    eErrCode   := E_DL_FlowMassConvErr.eInvalidUnit; // 故障级：目标单位越域 / Fault: destination out of domain
    RETURN;
END_CASE

(* —— 段 4：中介值与结果复检（四段式第四段） —— *)
IF (_fHub <> _fHub) OR ((_fHub - _fHub) <> DL_FMC_ZERO)
    OR (fConverted <> fConverted) OR ((fConverted - fConverted) <> DL_FMC_ZERO) THEN
    fConverted := DL_FMC_ZERO;                       // 复检异常回哨兵 / Recheck failed: sentinel
    eErrCode   := E_DL_FlowMassConvErr.eNonFinite;   // 故障级码 / Fault-level code
    RETURN;
END_IF

(* —— 段 5：成功出口（零值单列信息码） —— *)
IF (fValue < DL_FMC_EPS) AND (fValue > -DL_FMC_EPS) THEN
    eErrCode := E_DL_FlowMassConvErr.eZeroValue;     // 信息级：零流量 / Info: zero flow
ELSE
    eErrCode := E_DL_FlowMassConvErr.eOk;            // 信息级：换算完成 / Info: conversion completed
END_IF
FC_DL_FlowMassUnitConvert := TRUE;                   // 换算有效 / Conversion valid
END_FUNCTION

(* ---- FC_DL_FlowUnitConvert.st ---- *)
(*
  ==================================================================
  组件名 Component  : FC_DL_FlowUnitConvert
  分类   Category   : DL_MathData
  前缀   Naming     : FC_DL_ ｜ b/n/u/f/t/e/st 类型前缀制（R265）
  码位   Code ID    : 16#0001_0667（故障级）
  版本   Version    : 1.0.1
  复杂度 Complexity  : 低
  功能   Purpose    : 流量单位换算：m³/h ↔ L/min ↔ NL/min ↔ SCFM 四单位互转，
                      经 m³/h 基准单位两级换算；与 FC_DL_TempUnitConvert /
                      FC_DL_PressUnitConvert 同族三件齐（T0-4 单位换算族补口）。
  开源溯源 Origin    : T0-4 单位换算族补口（内部来源，零检索）；换算因子取
                      NIST 公开物理常数口径（1 ft³ = 0.0283168 m³，标准状态
                      60°F / 1 atm）；与 Temp / Press 族同骨架复用（本库自有
                      范式），零代码复制。
  许可证 License    : MIT
  参考   Reference  : IEC 61131-3:2013 §6.6 算术运算符；NIST 公开单位换算
                      常数口径
  平台   Platform   : 纯 IEC 61131-3（CASE / 四则），三平台通用
  依赖   Depends    : 无（零委托、零库件）
  分工声明 Split     : FC_DL_TempUnitConvert / FC_DL_PressUnitConvert 为同族
                      姊妹件（互引，三件齐口径）；本件只换流量，体积流量
                      与质量流量换算（需密度）归 FC_DL_FlowMassConvert
                      职责，本件不做（R216）。
  归属 Ownership     : E_DL_FlowUnit 属主为本文件（全库唯一定义，R264）；
                      引用件只引用不重声明。
  ------------------------------------------------------------------
  边界 Boundary     :
                      一 非有限闸：fValue 非有限（NaN / ±Inf）→ 故障级 0667 +
                         fResult = 0 + bValid = FALSE + 早退；
                      二 单位枚举闸：eUnitFrom / eUnitTo 任一越域（强改非法
                         枚举值）由 CASE ... ELSE 拦截 → 同码 0667 同形出口
                         （禁静默换算）；与非有限出口组合完全相同（fResult
                         = 0、bValid = FALSE、bError = TRUE），合并一码
                         （反证句见码表）；
                      三 换算链：fBase = fValue × 源因子（→ m³/h 基准），
                         fResult = fBase ÷ 目标因子；除子为目标因子常量
                         （因子表全部 > 0，编译期常量，除零不可达，R1 口径）；
                      四 负值合法（反向流量信号照实换算），零值合法；
                      五 NL/min 口径声明：标准状态取 0°C / 101.325 kPa，
                         1 NL/min = 0.06 m³/h；SCFM 取 60°F / 1 atm，
                         1 SCFM = 1.699011 m³/h（NIST 口径，常量注释逐条带
                         来源）；不同标准态需求由调用方先归一再入参；
                      六 纯函数：无记忆量、无定时器、无边沿实例，每调用重算；
                      七 无循环、无数组访问；无全局、无外部变量、无物理地址。
  错误码 Codes      :
    16#0001_0667【故障级】fValue 非有限或单位枚举越域（两场景出口同形，合并一码）
  码位反证 Note     :
    0667 合并「数值非有限」与「单位枚举越域」的理由：两场景出口组合完全相同
    （fResult = 0、bValid = FALSE、bError = TRUE），三组以内输出无法唯一还原
    该场景，按 R90 不另立码；非零正常换算无码。
  验收 Acceptance   :
    算法已证（脚本）：未跑 ｜ 编译器已证（三平台）：未跑
    V1 60 m³/h → L/min = 1000.0；V2 100 L/min → m³/h = 6.0
    V3 50 NL/min → m³/h = 3.0；V4 100 SCFM → m³/h ≈ 169.9011
    V5 同单位换算（eFrom = eTo）→ 原值返回（恒等链）
    V6 fValue = NaN → 码 0667 + fResult 0 + bValid = FALSE
    V7 eUnitFrom = 99（强改非法）→ 同码同形出口
    V8 负值 -6 m³/h → L/min = -100.0（反向流量照实）
  修订记录 Revision  :
    2026-11-21  v1.0.0  R64 首版（批 2 · 序号 6，T0-4 单位换算族补口，三件齐）
    2026-11-21  v1.0.1  R64 终审 R64-S1（严重·安全侧就地修）：DL_FUC_LMIN 因子
                       方向倒置（16.666667 为 [L/min 每 m³/h] 的倒数值，与本表
                       声明的 [（m³/h）/（L/min）] 口径相反）→ L/min 参与的全部
                       换算错 277.78 倍；改为 1 L/min = 0.06 m³/h。V1~V4 验收向量
                       修复后自证成立（V1 600000/0.06=1000.0 等），与 Press / Temp
                       姊妹件「因子 = 基准/源单位」口径统一。
  ==================================================================
*)
TYPE E_DL_FlowUnit :
(
    eM3h   := 0, // 立方米每小时 [m³/h]（基准单位）/ the cubic meter per hour, the canonical unit
    eLmin  := 1, // 升每分钟 [L/min] / the liter per minute
    eNLmin := 2, // 标准升每分钟 [NL/min]，0°C / 101.325 kPa / the normal liter per minute at the normal state
    eScfm  := 3  // 标准立方英尺每分钟 [SCFM]，60°F / 1 atm / the standard cubic foot per minute
);
END_TYPE

FUNCTION FC_DL_FlowUnitConvert : BOOL
VAR_INPUT
    fValue    : LREAL := 0.0;            // 入口流量值 [源单位]，必须有限 / the inlet flow value, must be finite
    eUnitFrom : E_DL_FlowUnit := E_DL_FlowUnit.eM3h;  // 源单位 [枚举] / the source unit
    eUnitTo   : E_DL_FlowUnit := E_DL_FlowUnit.eLmin;  // 目标单位 [枚举] / the target unit
END_VAR
VAR_OUTPUT
    fResult: LREAL; // 换算结果 [目标单位]，失败 = 0 / the converted result, zero on failure
    bValid : BOOL;  // 结果可用 [-] / the result usable flag
    eErr   : UDINT; // 错误码，0 = 正常 / the error code, zero is ok
    bError : BOOL;  // 故障标志（故障级码同拍置位，R45 配对）/ the fault flag raised with a fault level code
END_VAR
VAR
    fBase : LREAL := 0.0; // 基准量工作副本 [m³/h] / the canonical working copy in the cubic meter per hour
    fFromF: LREAL := 0.0; // 源单位因子 [（m³/h）/ 源单位] / the source unit factor to the canonical
    fToF  : LREAL := 0.0; // 目标单位因子 [（m³/h）/ 目标单位] / the target unit factor to the canonical
END_VAR  // R64 结构补齐：VAR 段缺失的 END_VAR（门禁机械修复）
VAR CONSTANT
    DL_FUC_ZERO   : LREAL := 0.0;      // 实数零常量 [目标单位] / the real zero constant
    DL_FUC_M3H    : LREAL := 1.0;      // m³/h 基准因子 [（m³/h）/（m³/h）] / the canonical factor of itself
    DL_FUC_LMIN   : LREAL := 0.06;     // L/min 因子：1 L/min = 0.06 m³/h（60/1000）[（m³/h）/（L/min）] / the liter per minute factor
    DL_FUC_NLMIN  : LREAL := 0.06;     // NL/min 因子：1 NL/min = 0.06 m³/h（0°C / 101.325 kPa）[（m³/h）/（NL/min）] / the normal liter factor
    DL_FUC_SCFM   : LREAL := 1.699011; // SCFM 因子：1 SCFM = 0.0283168 × 60 m³/h（60°F / 1 atm，NIST 口径）[（m³/h）/（SCFM）] / the standard cubic foot factor
END_VAR

// 段 1｜返回值与全部出口预置安全值（R45 四段式第一段）/ segment 1, the preset of the return and all outlets
FC_DL_FlowUnitConvert := FALSE; // 返回值预置假 / preset the return false
fResult := DL_FUC_ZERO; // 结果预置零 [目标单位] / preset the result zero
bValid := FALSE; // 可用标志预置假 / preset the validity false
eErr := 16#0000_0000; // 错误码预置正常 / preset the code to ok
bError := FALSE; // 故障标志预置假 / preset the fault flag false
fBase := DL_FUC_ZERO; // 基准量预置零 [m³/h] / preset the canonical copy zero
fFromF := DL_FUC_M3H; // 源因子预置基准因子（ELSE 兜底口径）/ preset the source factor to the canonical
fToF := DL_FUC_M3H; // 目标因子预置基准因子（ELSE 兜底口径）/ preset the target factor to the canonical

// 段 2｜非有限闸（边界一）/ segment 2, the finiteness gate
IF (fValue <> fValue) OR ((fValue - fValue) <> (fValue - fValue)) THEN // 入口值非有限（NaN 或 ±Inf）/ the inlet value is not finite
    eErr := 16#0001_0667; // 故障级：非有限或单位越域（合并一码，R90）/ fault grade under the merged code
    bError := TRUE; // 同拍置故障标志（R45 配对）/ raise the fault flag on the same scan
    bValid := FALSE; // 结果不可用 / the result is not usable
    RETURN; // 早退 / early return
END_IF

// 段 3｜源单位因子表（边界二：CASE ... ELSE 拦非法枚举）/ segment 3, the source factor table with the illegal guard
CASE eUnitFrom OF
    E_DL_FlowUnit.eM3h:   fFromF := DL_FUC_M3H;   // 基准因子 / the canonical factor
    E_DL_FlowUnit.eLmin:  fFromF := DL_FUC_LMIN;  // L/min 因子 / the liter per minute factor
    E_DL_FlowUnit.eNLmin: fFromF := DL_FUC_NLMIN; // NL/min 因子 / the normal liter factor
    E_DL_FlowUnit.eScfm:  fFromF := DL_FUC_SCFM;  // SCFM 因子 / the standard cubic foot factor
    ELSE // 非法枚举拦截（禁静默换算，边界二）/ the illegal enumeration guard
        eErr := 16#0001_0667; // 故障级：单位越域（与非有限同形出口，R90）/ fault grade, the unit out of the domain
        bError := TRUE; // 同拍置故障标志（R45 配对）/ raise the fault flag on the same scan
        bValid := FALSE; // 结果不可用 / the result is not usable
        RETURN; // 早退 / early return
END_CASE

// 段 4｜目标单位因子表（边界二：CASE ... ELSE 拦非法枚举）/ segment 4, the target factor table with the illegal guard
CASE eUnitTo OF
    E_DL_FlowUnit.eM3h:   fToF := DL_FUC_M3H;   // 基准因子 / the canonical factor
    E_DL_FlowUnit.eLmin:  fToF := DL_FUC_LMIN;  // L/min 因子 / the liter per minute factor
    E_DL_FlowUnit.eNLmin: fToF := DL_FUC_NLMIN; // NL/min 因子 / the normal liter factor
    E_DL_FlowUnit.eScfm:  fToF := DL_FUC_SCFM;  // SCFM 因子 / the standard cubic foot factor
    ELSE // 非法枚举拦截（禁静默换算，边界二）/ the illegal enumeration guard
        eErr := 16#0001_0667; // 故障级：单位越域（与非有限同形出口，R90）/ fault grade, the unit out of the domain
        bError := TRUE; // 同拍置故障标志（R45 配对）/ raise the fault flag on the same scan
        bValid := FALSE; // 结果不可用 / the result is not usable
        RETURN; // 早退 / early return
END_CASE

// 段 5｜两级换算（边界三：除子 fToF 为常量因子，因子表全部 > 0，除零不可达）/ segment 5, the two stage conversion with the proven constant divisor
fBase := fValue * fFromF; // 源单位 → m³/h 基准 [m³/h] / the source value to the canonical
fResult := fBase / fToF; // 基准 → 目标单位 [目标单位]（除子常量已证 > 0）/ the canonical to the target with the proven divisor
bValid := TRUE; // 结果可用 / the result is usable
FC_DL_FlowUnitConvert := TRUE; // 返回成功 / return success
END_FUNCTION

(* ---- FC_DL_ForceUnitConvert.st ---- *)
(*==============================================================================
 * 组件名称 : FC_DL_ForceUnitConvert ｜ 子库 : DL_MathData ｜ v1.0.0 ｜ 2026-11-23
 * 平台     : CODESYS 3.5 / TwinCAT 3 / InoProShop / Machine Expert（纯 IEC，无厂商库）
 * 功能简介 : 力单位 N / kN / lbf（磅力）两两互转。源/目标由枚举对单向选择，
 *            单向基准链（先归一到 N）使公式域固定为 3+3 条分支。
 * 契约     : 返回换算结果 [目标单位]；枚举非法（越界值）返回 0.0；
 *            除数为编译期非零常量，无除零风险；纯函数无状态。
 * 依赖     : 无 DL_ 内部依赖（本批自足实现）
 * 红线自检 : R1 零全局 R2 零%I/%Q R3 纯IEC R4 枚举越界拒收返 0 + 常量除数
 *            R5 全变量与枚举项双语同行注释 R6 N/A（无状态机） R7 N/A
 * 修订历史 : 2026-11-23 R78-B1 工程单位换算族模板派生首版
 *============================================================================*)
TYPE E_DL_ForceUnit :
(
    eN := 0,        // 牛顿 [N] / Newton
    eKN,            // 千牛 [kN] / Kilo-newton
    eLbf            // 磅力 [lbf] / Pound-force
);
END_TYPE

FUNCTION FC_DL_ForceUnitConvert : REAL
VAR_INPUT
    fValue : REAL;          // 输入数值 [源单位] / Input value in source unit
    eSrc : E_DL_ForceUnit;  // 源单位选择 / Source unit selector
    eDst : E_DL_ForceUnit;  // 目标单位选择 / Destination unit selector
END_VAR
VAR
    fBase : REAL;           // 归一化中间值 [N] / Normalized intermediate in newtons
END_VAR
FC_DL_ForceUnitConvert := 0.0;  // 缺省返回 0 / Default return 0
CASE eSrc OF                    // 段 1：归一到基准 N / Normalize to base newtons
    E_DL_ForceUnit.eN: fBase := fValue;                     // 基准直通 / Base pass-through
    E_DL_ForceUnit.eKN: fBase := fValue * 1000.0;           // 1 kN = 1000 N
    E_DL_ForceUnit.eLbf: fBase := fValue * 4.4482216;       // 1 lbf = 4.4482216 N（公开定义）
    ELSE FC_DL_ForceUnitConvert := 0.0; RETURN;             // 源枚举非法返 0 / Invalid source returns 0
END_CASE
CASE eDst OF                    // 段 2：基准到目标 / Base to destination
    E_DL_ForceUnit.eN: FC_DL_ForceUnitConvert := fBase;                 // 基准直通 / Base pass-through
    E_DL_ForceUnit.eKN: FC_DL_ForceUnitConvert := fBase / 1000.0;       // N 到 kN
    E_DL_ForceUnit.eLbf: FC_DL_ForceUnitConvert := fBase / 4.4482216;   // N 到 lbf
    ELSE FC_DL_ForceUnitConvert := 0.0;                     // 目标枚举非法返 0 / Invalid destination returns 0
END_CASE
END_FUNCTION

(* ---- FC_DL_HarmonicSpectrumBin.st ---- *)
(*
  FC_DL_HarmonicSpectrumBin  —  单频点 DFT 幅值·相位提取 / Single-bin DFT magnitude and phase extraction
  分类 Category : DL_MathData
  码位 Code     : 16#05_0_00
  版本 Version  : 1.0.0
  来源标签 Tag  : t2-1-lgf-math
  溯源 Source   : LGF Math 语义借鉴 · clean-room 实现，仅借分类/参数域/命名，未复制源码行
  功能 Function : 1) Goertzel 递推单频点 DFT，矩形/Hann 双窗，Hann 相干增益 0.5 做幅值修正；
                  2) 相位解卷并给贴轴归属（imag = 0 且 real < 0 归正支，返回域 (-180, 180] 度）；
                  3) 五道边界闸：窗长域 / 采样率 / 奈奎斯特 / 窗内非有限样本 / 幅值分辨力下限。
  边界 Boundary : ① nWindowSize 越 [8, 1023] 判无效置故障码，不进入循环；
                  ② fSampleRateHz <= 0 先判零再除（防除零），判零前先过非有限闸；
                  ③ fTargetFreqHz >= 奈奎斯特判无效，宁可不报也不混叠出假值；
                  ④ 窗内任一 NaN/Inf 整窗无效（自反判 NaN + 差值自减判 Inf 双判）；
                  ⑤ 幅值 < fMagFloor 输出 0 并置信息码，不置 bError。
  依赖 Depends  : FC_DL_NthRoot（开方 nRoot = 2；本件禁内联 SQRT 原语，R140 委托优先）
  纯函数声明    : 本件为纯函数，零内部状态、零跨周期驻留、零 GVL/物理地址引用

  码表 Error codes（本件格 05_0_00，子码步进 +0x10）:
    16#0005_0500 故障级：组态非法（窗长越域 / 采样率 <= 0 / 目标频率 >= 奈奎斯特 / 幅值门限 < 0 / 组态量非有限）
    16#0005_0510 信息级：窗内存在非有限样本整窗无效 / 幅值低于分辨力（不置 bError）

  修订历史 Revision :
    2026-11-18  v1.0.0  R36 首版入库（W1 窗首件）
*)

TYPE E_DL_SpectrumWindow :
(
    eRect := 0,   // 矩形窗，相干增益 1.0（频率分辨率最优，泄漏最大）/ Rectangular window, coherent gain 1.0
    eHann := 1    // Hann 窗，相干增益 0.5（抑制泄漏）/ Hann window, coherent gain 0.5
);
END_TYPE

FUNCTION FC_DL_HarmonicSpectrumBin : BOOL
VAR_INPUT
    afSampleBuffer : ARRAY[0..1023] OF LREAL;                  // 采样窗缓冲区，索引 0 为最早样本 / Sample window buffer, index 0 = oldest sample
    nWindowSize    : UINT := 0;                                // 有效窗长 [样本数]，域 8 ~ 1023 / Effective window length [samples]
    fSampleRateHz  : LREAL := 0.0;                             // 采样率 [Hz]，域 > 0 / Sampling rate [Hz], domain > 0
    fTargetFreqHz  : LREAL := 0.0;                             // 目标提取频率 [Hz]，域 [0, 奈奎斯特) / Target bin frequency [Hz]
    fMagFloor      : LREAL := 1.0E-6;                          // 幅值分辨力下限 [输入物理量单位]，域 >= 0 / Magnitude floor [EU]
    eWindowType    : E_DL_SpectrumWindow := E_DL_SpectrumWindow.eRect; // 窗型选择 / Window type selection
END_VAR
VAR_OUTPUT
    fMagnitude : LREAL;                                        // 峰值幅值输出，物理量单位随输入 [EU] / Peak magnitude [EU]
    fPhaseDeg  : LREAL;                                        // 相位输出 [deg]，域 (-180, 180] / Phase [deg]
    bValid     : BOOL;                                         // 结果有效标志，FALSE 时幅值相位均为 0 / Result valid flag
    bError     : BOOL;                                         // 故障标志，与故障级码配对 / Fault flag paired with fault code
    nErrId     : UDINT;                                        // 事件码，0 = 无事件 / Event code, 0 = no event
END_VAR
VAR
    nIdx          : INT;                                       // 样本循环索引 [1] / Sample loop index
    nCount        : INT;                                       // 生效窗长整型副本 [样本数] / Integer copy of window length
    fOmega        : LREAL;                                     // 数字角频率 [rad] / Digital angular frequency [rad]
    fCoeff        : LREAL;                                     // Goertzel 递推系数 2·cos(ω) [1] / Goertzel recursion coefficient
    fS0           : LREAL;                                     // 递推当前拍状态量 [EU] / Recursion state, current
    fS1           : LREAL;                                     // 递推前一拍状态量 [EU] / Recursion state, previous
    fS2           : LREAL;                                     // 递推前二拍状态量 [EU] / Recursion state, two scans back
    fWin          : LREAL;                                     // 当前样本窗权值 [1] / Window weight of current sample
    fCoherentGain : LREAL;                                     // 窗相干增益 [1]，矩形 1.0 / Hann 0.5 / Coherent gain of window
    fSample       : LREAL;                                     // 当前样本值副本 [EU] / Copy of current sample
    fPower        : LREAL;                                     // Goertzel 功率量（未开方）[EU^2] / Goertzel power term
    fMagRaw       : LREAL;                                     // 窗修正前幅值 [EU] / Magnitude before window correction
    fReal         : LREAL;                                     // 相位实部（s1 - s2·cosω）[EU] / Phase real part
    fImag         : LREAL;                                     // 相位虚部（s2·sinω）[EU] / Phase imaginary part
    fPhaseRad     : LREAL;                                     // 相位弧度中间量 [rad] / Phase in radians
    fNyquist      : LREAL;                                     // 奈奎斯特频率 fSampleRateHz / 2 [Hz] / Nyquist frequency [Hz]
    bNonFinite    : BOOL;                                      // 窗内非有限样本标志 / Non-finite sample flag
    bSqrtValid    : BOOL;                                      // 开方委托结果有效标志 / Sqrt delegation valid flag
    fSqrtOut      : LREAL;                                     // 开方委托返回值 [EU] / Sqrt delegation return value
END_VAR
VAR CONSTANT
    DL_WIN_MIN  : UINT  := 8;                      // 窗长下限 [样本数]，低于此值分辨率无工程意义 / Window length lower bound
    DL_WIN_MAX  : UINT  := 1023;                   // 窗长上限 [样本数]，等于缓冲区上界 / Window length upper bound
    DL_TWO_PI   : LREAL := 6.283185307179586477;   // 2π LREAL 精度字面量 [rad] / 2π in LREAL precision
    DL_RAD2DEG  : LREAL := 57.295779513082320877;  // 弧度转度 [deg/rad] / Radian to degree factor
    DL_EPS      : LREAL := 1.0E-12;                // 判零容差 [1] / Zero tolerance
END_VAR

(* —— 段 0：返回值与输出预置安全值（纯函数，无状态刷新） —— *)
FC_DL_HarmonicSpectrumBin := FALSE;   // 返回布尔：FALSE = 本拍无有效结果
fMagnitude   := 0.0;                  // 幅值预置 0 [EU]
fPhaseDeg    := 0.0;                  // 相位预置 0 [deg]
bValid       := FALSE;                // 有效标志预置 FALSE
bError       := FALSE;                // 故障标志预置 FALSE（故障级码赋值后 3 行内置位）
nErrId       := 0;                    // 事件码预置 0
nCount       := UINT_TO_INT(nWindowSize);  // 窗长整型副本 [样本数]
fCoherentGain := 1.0;                 // 相干增益默认矩形窗 [1]
bNonFinite   := FALSE;                // 非有限标志预置 FALSE
fNyquist     := fSampleRateHz * 0.5;  // 奈奎斯特频率 [Hz]，采样率闸命中前仅作占位

(* —— 段 1：组态域闸（R151 覆盖全部参与换算的引脚） —— *)
IF (fSampleRateHz <> fSampleRateHz) OR ((fSampleRateHz - fSampleRateHz) <> (fSampleRateHz - fSampleRateHz)) THEN
    nErrId := 16#0005_0500;           // 故障级：采样率非有限（NaN 自反 / Inf 差值自减）
    bError := TRUE;                   // 故障标志置位（R45 配对）
    RETURN;                           // 域闸命中不调内核
END_IF
IF (fTargetFreqHz <> fTargetFreqHz) OR ((fTargetFreqHz - fTargetFreqHz) <> (fTargetFreqHz - fTargetFreqHz)) THEN
    nErrId := 16#0005_0500;           // 故障级：目标频率非有限
    bError := TRUE;                   // 故障标志置位（R45 配对）
    RETURN;                           // 域闸命中不调内核
END_IF
IF (fMagFloor <> fMagFloor) OR (fMagFloor < 0.0) THEN
    nErrId := 16#0005_0500;           // 故障级：幅值门限非有限或为负
    bError := TRUE;                   // 故障标志置位（R45 配对）
    RETURN;                           // 域闸命中不调内核
END_IF
IF (nWindowSize < DL_WIN_MIN) OR (nWindowSize > DL_WIN_MAX) THEN
    nErrId := 16#0005_0500;           // 故障级：窗长越 [8, 1023] 域（下界防退化，上界防数组越界）
    bError := TRUE;                   // 故障标志置位（R45 配对）
    RETURN;                           // 不进入循环
END_IF
IF fSampleRateHz <= 0.0 THEN
    nErrId := 16#0005_0500;           // 故障级：采样率 <= 0（除零前置判定）
    bError := TRUE;                   // 故障标志置位（R45 配对）
    RETURN;                           // 域闸命中不调内核
END_IF
IF (fTargetFreqHz < 0.0) OR (fTargetFreqHz >= fNyquist) THEN
    nErrId := 16#0005_0500;           // 故障级：目标频率越 [0, 奈奎斯特) 域，拒绝混叠假值
    bError := TRUE;                   // 故障标志置位（R45 配对）
    RETURN;                           // 域闸命中不调内核
END_IF

(* —— 段 2：内核参数（角频率与递推系数），窗型决定相干增益 —— *)
fOmega := DL_TWO_PI * fTargetFreqHz / fSampleRateHz;   // 数字角频率 [rad]，采样率已证明 > 0
fCoeff := 2.0 * COS(fOmega);                           // 递推系数 [1]
IF eWindowType = E_DL_SpectrumWindow.eHann THEN
    fCoherentGain := 0.5;                              // Hann 窗相干增益 [1]
ELSE
    fCoherentGain := 1.0;                              // 矩形窗（含未知枚举值兜底）相干增益 [1]
END_IF

(* —— 段 3：Goertzel 递推主循环（样本数已钳在数组域内，循环计数器结构上有界） —— *)
fS1 := 0.0;                                            // 递推状态清零
fS2 := 0.0;                                            // 递推状态清零
FOR nIdx := 0 TO (nCount - 1) DO
    fSample := afSampleBuffer[nIdx];                   // 取样本 [EU]
    IF (fSample <> fSample) OR ((fSample - fSample) <> (fSample - fSample)) THEN
        bNonFinite := TRUE;                            // 窗内出现 NaN 或 Inf
    END_IF
    IF eWindowType = E_DL_SpectrumWindow.eHann THEN
        fWin := 0.5 - 0.5 * COS(DL_TWO_PI * INT_TO_LREAL(nIdx) / INT_TO_LREAL(nCount - 1));  // Hann 窗权值 [1]
    ELSE
        fWin := 1.0;                                   // 矩形窗权值 [1]
    END_IF
    fS0 := fWin * fSample + fCoeff * fS1 - fS2;         // 递推当前拍 [EU]
    fS2 := fS1;                                         // 状态后移
    fS1 := fS0;                                         // 状态后移
END_FOR

IF bNonFinite THEN
    nErrId := 16#0005_0510;           // 信息级：窗内非有限样本，整窗无效（信息级不置 bError）
    RETURN;                           // 不出结论
END_IF

(* —— 段 4：功率量 → 幅值（委托 FC_DL_NthRoot 开方，禁内联 SQRT），相位解卷 —— *)
fPower := fS1 * fS1 + fS2 * fS2 - fCoeff * fS1 * fS2;   // Goertzel 功率量 [EU^2]
IF fPower < 0.0 THEN
    fPower := 0.0;                                      // 数值负偏钳零（不动点舍入噪声）
END_IF
fSqrtOut := FC_DL_NthRoot(fValue := fPower, nRoot := 2, bValid => bSqrtValid);  // 委托开方
IF NOT bSqrtValid THEN
    nErrId := 16#0005_0510;           // 信息级：开方委托判无效（功率量非有限）
    RETURN;                           // 不出结论
END_IF
fMagRaw := 2.0 * fSqrtOut / INT_TO_LREAL(nCount);                        // 单边幅值（未做窗修正）[EU]
fMagnitude := fMagRaw / fCoherentGain;                                    // 窗相干增益修正后幅值 [EU]
IF (fMagnitude <> fMagnitude) OR ((fMagnitude - fMagnitude) <> (fMagnitude - fMagnitude)) THEN
    fMagnitude := 0.0;                                                    // 非有限复检兜底
    nErrId := 16#0005_0510;           // 信息级：幅值非有限
    RETURN;                           // 不出结论
END_IF

fReal := fS1 - fS2 * COS(fOmega);                       // 相位实部 [EU]
fImag := fS2 * SIN(fOmega);                             // 相位虚部 [EU]
IF (ABS(fReal) < DL_EPS) AND (ABS(fImag) < DL_EPS) THEN
    fPhaseRad := 0.0;                                   // 零幅（数值退化）相位无意义，取 0
ELSIF fImag >= 0.0 THEN
    fPhaseRad := ATAN(fImag / (ABS(fReal) + DL_EPS));    // 上支（含 imag = 0 且 real < 0）[rad]
    IF fReal < 0.0 THEN
        fPhaseRad := fPhaseRad + DL_TWO_PI * 0.5;       // 第二象限贴轴归属到正支 [rad]
    END_IF
ELSE
    fPhaseRad := ATAN(fImag / (ABS(fReal) + DL_EPS));    // 下支 [rad]
    IF fReal < 0.0 THEN
        fPhaseRad := fPhaseRad - DL_TWO_PI * 0.5;       // 第三象限贴轴归属到负支 [rad]
    END_IF
END_IF
fPhaseDeg := fPhaseRad * DL_RAD2DEG;                    // 相位 [deg]，域 (-180, 180]

(* —— 段 5：分辨力下限判定（低幅不出结论，置信息码） —— *)
IF fMagnitude < fMagFloor THEN
    fMagnitude := 0.0;                // 低于分辨力输出 0 [EU]
    nErrId := 16#0005_0510;           // 信息级：幅值低于分辨力（信息级不置 bError）
    RETURN;                           // 不出结论
END_IF

bValid := TRUE;                       // 结果有效
FC_DL_HarmonicSpectrumBin := TRUE;    // 返回布尔：TRUE = 本拍有有效结果

END_FUNCTION

(* ---- FC_DL_HumidityUnitConvert.st ---- *)
(*==============================================================================
 * 组件名称 (Component)  : FC_DL_HumidityUnitConvert
 * 所属子库 (Sublibrary) : DL_MathData
 * 当前版本 (Version)    : 1.0.0
 * 兼容性   (Platform)   : CODESYS 3.5+ / TwinCAT 3 / 汇川 InoProShop / 施耐德 Machine Expert
 *                         仅依赖 IEC 61131-3 标准数学（EXP），零厂商私有库
 * 功能描述 (Function)   : 湿度换算：相对湿度 RH% ↔ 绝对湿度 AH[g/m³]。
 *                         饱和水汽压用 Magnus 近似式（WMO 常用系数）：
 *                           Psat(T) = 6.112 × EXP(17.62 × T / (243.12 + T))    [hPa]
 *                           AH = (RH/100) × 216.7 × Psat(T) / (T + 273.15)    [g/m3]
 *                           RH = AH × (T + 273.15) / (216.7 × Psat(T)) × 100  [%]
 *                         两式互为反函数（AH 侧以 fValue 为 AH 求 RH，反之亦然），
 *                         故本件自成闭环，不依赖外部湿度表。
 * 接口     (Interface)  : 输入 fValue 被换算湿度 [源单位]、eSrc 源单位、eDst 目标单位、
 *                         fTempC 干球温度 [℃]（**换算必需，非可选**）；
 *                         输出 fConverted 换算结果 [目标单位]、eErrCode（E_DL_HumConvErr）；
 *                         返回值 = bValid 数值可信标志（TRUE = fConverted 可信）。
 * 边界     (Boundary)   : ① 属主边界：只做 RH↔AH 换算，不做露点 / 焓值 / 湿球温度计算。
 *                         ② **适用域**：干球温度 -40..80 ℃（Magnus 式标定域），超域 → 故障级
 *                         eTempOutOfRange（外推会显著失真，禁止静默外推）。
 *                         ③ **全部浮点入参做非有限双判**（fValue 与 fTempC 逐一枚举，
 *                         含换算用的温度量，防止 NaN 温度使结果静默失效）。
 *                         ④ RH 源值域 0..100，超域 → 故障级 eRhOutOfRange。
 *                         AH 源值必须非负，负值 → 故障级 eNegativeValue。
 *                         ⑤ 反算 RH 结果超 100（过饱和）→ 钳位 100 并置信息级 eClampRh。
 *                         ⑥ 分母防护：Psat 恒 > 0（指数函数）；(243.12+T) 在适用域内恒 >= 203.12；
 *                         (T+273.15) 在适用域内恒 >= 233.15；另加显式判零分支作双保险。
 *                         ⑦ 零全局耦合（无 GVL / VAR_EXTERNAL / 物理地址）。
 * 分工声明 (Scope)      : 与 `FC_DL_ConcentrationUnitConvert` 分工：气体浓度归那件；
 *                         与露点/焓值件（未入库）分工：本件不含相变焓计算。
 * 来源标签 (Source Tag) : 开源溯源：lgf-math 换算系数（公开物理常数，clean-room 重写）；许可证 MIT（仅参考语义，代码原创）
 * 码表     (Codes)      : 本件不占用全局数字码位；出口为 BOOL + LREAL +
 *                         本文件内定义 enum E_DL_HumConvErr（全库唯一）。
 * 红线自检 (Redline)    : R1 ✓ 零 GVL/VAR_EXTERNAL ｜ R2 ✓ 零 %I/%Q/%M ｜ R3 ✓ 纯 IEC 61131-3
 *                         R4 ✓ 全部浮点入参非有限双判 + 温度域闸 + RH 域闸 + 分母显式判零 ｜ R5 ✓ 声明逐行同行双语注释
 *                         R6 N/A（纯函数无状态机） ｜ R7 N/A（无实例调用）
 * 修订历史 (Revision)   : 2026-11-23  v1.0.0  R77 首版（批次 B2 · 序号 19）
 * 验收向量 (Acceptance) : ① fValue=50.0(RH), eSrc=eRhPercent, eDst=eAbsGm3, fTempC=25.0 →
 *                         Psat=6.112×EXP(17.62×25/268.12)=31.6713 hPa（容差 1E-3），
 *                         AH=0.5×216.7×31.6713/298.15 ≈ 11.511 g/m3（容差 1E-2）；
 *                         ② fValue=11.511, eSrc=eAbsGm3, eDst=eRhPercent, fTempC=25.0 →
 *                         RH ≈ 50.0 %（容差 1E-2，与 ① 互逆）；
 *                         ③ eSrc=eDst 直通：fValue=42.0 原样返回，eOk；
 *                         ④ fTempC=100.0 → 返回 FALSE, 0, eTempOutOfRange；
 *                         ⑤ fValue=120.0(RH), eSrc=eRhPercent → 返回 FALSE, 0, eRhOutOfRange。
 *==============================================================================*)

(*-----------------------------------------------------------------------------
 * 枚举: E_DL_HumUnit（湿度单位表，归属 DL_MathData，与本件同文件，全库唯一属主）
 *----------------------------------------------------------------------------*)
TYPE E_DL_HumUnit :
(
    eRhPercent := 0,   // 相对湿度（百分数） [%RH] / Relative humidity in percent
    eAbsGm3    := 1    // 绝对湿度（每立方米水汽克数） [g/m3] / Absolute humidity in grams per cubic metre
);
END_TYPE

(*-----------------------------------------------------------------------------
 * 枚举: E_DL_HumConvErr（湿度换算错误码）
 *----------------------------------------------------------------------------*)
TYPE E_DL_HumConvErr :
(
    eOk             := 0,   // 信息级：换算完成 / Info: conversion completed
    eClampRh        := 1,   // 信息级：反算 RH 过饱和已钳位 100 / Info: computed RH clamped to 100
    eInvalidUnit    := 2,   // 故障级：单位枚举越域 / Fault: unit enum out of domain
    eNonFinite      := 3,   // 故障级：入参非有限 / Fault: non-finite input
    eTempOutOfRange := 4,   // 故障级：干球温度超出 Magnus 标定域 / Fault: dry-bulb temperature out of calibrated range
    eRhOutOfRange   := 5,   // 故障级：RH 源值超出 0..100 / Fault: RH source out of range
    eNegativeValue  := 6    // 故障级：AH 源值为负 / Fault: negative absolute humidity
);
END_TYPE

FUNCTION FC_DL_HumidityUnitConvert : BOOL
VAR_INPUT
    fValue : LREAL;         // 被换算湿度值 [源单位] / Humidity value in source unit
    eSrc   : E_DL_HumUnit;  // 源单位枚举 [-] / Source unit enum
    eDst   : E_DL_HumUnit;  // 目标单位枚举 [-] / Destination unit enum
    fTempC : LREAL;         // 干球温度（换算必需） [℃] / Dry-bulb temperature, mandatory for conversion [degC]
END_VAR
VAR_OUTPUT
    fConverted : LREAL;           // 换算结果 [目标单位] / Converted result
    fSatPress  : LREAL;           // 饱和水汽压（诊断用） [hPa] / Saturation vapour pressure, diagnostic [hPa]
    eErrCode   : E_DL_HumConvErr; // 错误码出口 [-] / Error code outlet
END_VAR
VAR
    _bNonFin : BOOL;   // 入参非有限当拍标志 [-] / Non-finite input flag
    _fDen    : LREAL;  // 显式分母防护量 [-] / Explicit denominator guard value
    _fRat    : LREAL;  // 中间比值（RH 分数 / 缩放后 AH） [-] / Intermediate ratio
END_VAR
VAR CONSTANT
    DL_HUC_A     : LREAL := 17.62;     // Magnus 分子系数 [-] / Magnus numerator coefficient
    DL_HUC_B     : LREAL := 243.12;    // Magnus 分母常数 [℃] / Magnus denominator constant
    DL_HUC_C     : LREAL := 6.112;     // 0 ℃ 饱和水汽压 [hPa] / Saturation pressure at zero degC
    DL_HUC_K     : LREAL := 216.7;     // 水汽气体常数换算因子 [g/m3 per hPa] / Water vapour conversion factor
    DL_HUC_KABS  : LREAL := 273.15;    // 摄氏转开尔文偏移 [K] / Celsius to Kelvin offset
    DL_HUC_HUND  : LREAL := 100.0;     // 百分数换算因子 [-] / Percent scaling factor
    DL_HUC_TMIN  : LREAL := -40.0;     // 干球温度下限 [℃] / Dry-bulb lower bound [degC]
    DL_HUC_TMAX  : LREAL := 80.0;      // 干球温度上限 [℃] / Dry-bulb upper bound [degC]
    DL_HUC_RHMAX : LREAL := 100.0;     // 相对湿度上限 [%RH] / Relative humidity ceiling
    DL_HUC_ZERO  : LREAL := 0.0;       // 零基准与非有限判零基准 [-] / Zero and non-finite base
    DL_HUC_TINY  : LREAL := 1.0E-9;    // 分母近似零阈值 [-] / Near-zero denominator threshold
END_VAR

(* —— 段 0：出口预置安全值 —— *)
FC_DL_HumidityUnitConvert := FALSE;                // 返回值预置无效 / Return preset invalid
fConverted := DL_HUC_ZERO;                         // 结果哨兵 0 / Result sentinel
fSatPress  := DL_HUC_ZERO;                         // 饱和压哨兵 0 / Saturation pressure sentinel
eErrCode   := E_DL_HumConvErr.eInvalidUnit;        // 预置最严码 / Preset strictest code

(* —— 段 1：非有限域闸（每个浮点入参逐一枚举：湿度值与温度值） —— *)
_bNonFin := (fValue <> fValue) OR ((fValue - fValue) <> DL_HUC_ZERO);      // 湿度值非有限 / Humidity non-finite
_bNonFin := _bNonFin OR (fTempC <> fTempC) OR ((fTempC - fTempC) <> DL_HUC_ZERO);  // 温度值非有限 / Temperature non-finite
IF _bNonFin THEN
    eErrCode := E_DL_HumConvErr.eNonFinite;        // 故障级码 / Fault-level code
    RETURN;
END_IF

(* —— 段 2：干球温度域闸（Magnus 标定域，禁止外推） —— *)
IF (fTempC < DL_HUC_TMIN) OR (fTempC > DL_HUC_TMAX) THEN
    eErrCode := E_DL_HumConvErr.eTempOutOfRange;   // 故障级码 / Fault-level code
    RETURN;
END_IF

(* —— 段 3：单位枚举域闸（两侧成员逐一比较） —— *)
IF (eSrc <> E_DL_HumUnit.eRhPercent) AND (eSrc <> E_DL_HumUnit.eAbsGm3) THEN
    RETURN;                                        // 源单位越域：保持预置故障码 / Source unit out of domain
END_IF
IF (eDst <> E_DL_HumUnit.eRhPercent) AND (eDst <> E_DL_HumUnit.eAbsGm3) THEN
    RETURN;                                        // 目标单位越域：保持预置故障码 / Destination unit out of domain
END_IF

(* —— 段 4：饱和水汽压计算（分母 243.12+T 在适用域内 >= 203.12，仍显式判零） —— *)
_fDen := DL_HUC_B + fTempC;                        // Magnus 分母 / Magnus denominator
IF _fDen < DL_HUC_TINY THEN
    eErrCode := E_DL_HumConvErr.eTempOutOfRange;   // 分母异常：判温度越域 / Abnormal denominator: treat as out of range
    RETURN;
END_IF
fSatPress := DL_HUC_C * EXP(DL_HUC_A * fTempC / _fDen);   // 饱和水汽压 [hPa] / Saturation vapour pressure

(* —— 段 5：源值域闸（RH 侧 0..100，AH 侧非负） —— *)
IF eSrc = E_DL_HumUnit.eRhPercent THEN
    IF (fValue < DL_HUC_ZERO) OR (fValue > DL_HUC_RHMAX) THEN
        eErrCode := E_DL_HumConvErr.eRhOutOfRange; // 故障级：RH 越域 / Fault: RH out of range
        RETURN;
    END_IF
ELSE
    IF fValue < DL_HUC_ZERO THEN
        eErrCode := E_DL_HumConvErr.eNegativeValue; // 故障级：AH 为负 / Fault: negative absolute humidity
        RETURN;
    END_IF
END_IF

(* —— 段 6：换算主分支 —— *)
IF eSrc = eDst THEN
    fConverted := fValue;                          // 同单位直通，无舍入 / Same unit pass-through without rounding
    eErrCode   := E_DL_HumConvErr.eOk;             // 信息级成功 / Info success
ELSIF (eSrc = E_DL_HumUnit.eRhPercent) AND (eDst = E_DL_HumUnit.eAbsGm3) THEN
    _fRat := fValue / DL_HUC_HUND;                 // RH 化分数 / RH to fraction
    _fDen := fTempC + DL_HUC_KABS;                 // 绝对温标 / Absolute temperature
    IF _fDen < DL_HUC_TINY THEN
        eErrCode := E_DL_HumConvErr.eTempOutOfRange;  // 分母异常防护 / Denominator guard
        RETURN;
    END_IF
    fConverted := _fRat * DL_HUC_K * fSatPress / _fDen;   // AH = (RH/100)*216.7*Psat/(T+273.15)
    eErrCode   := E_DL_HumConvErr.eOk;             // 信息级成功 / Info success
ELSE
    (* AH → RH：分母 = 216.7 × Psat，Psat 恒正，仍显式判零作双保险 *)
    _fDen := DL_HUC_K * fSatPress;                 // 分母：水汽因子 × 饱和压 / Denominator: factor times saturation pressure
    IF _fDen < DL_HUC_TINY THEN
        eErrCode := E_DL_HumConvErr.eTempOutOfRange;  // 分母近似零防护 / Near-zero denominator guard
        RETURN;
    END_IF
    _fRat      := fValue * (fTempC + DL_HUC_KABS) / _fDen;   // AH × (T+273.15) / (216.7×Psat)
    fConverted := _fRat * DL_HUC_HUND;             // 化百分数 / Scale to percent
    IF fConverted > DL_HUC_RHMAX THEN
        fConverted := DL_HUC_RHMAX;                // 过饱和钳位 100 / Clamp supersaturation to 100
        eErrCode   := E_DL_HumConvErr.eClampRh;    // 信息级钳位码 / Info clamp code
    ELSE
        eErrCode   := E_DL_HumConvErr.eOk;         // 信息级成功 / Info success
    END_IF
END_IF

(* —— 段 7：结果非有限复检兜底（含饱和压复检） —— *)
IF (fConverted <> fConverted) OR ((fConverted - fConverted) <> DL_HUC_ZERO) THEN
    fConverted := DL_HUC_ZERO;                     // 复检异常回哨兵 / Recheck failed: sentinel
    eErrCode   := E_DL_HumConvErr.eNonFinite;      // 故障级码 / Fault-level code
    RETURN;
END_IF
IF (fSatPress <> fSatPress) OR ((fSatPress - fSatPress) <> DL_HUC_ZERO) OR (fSatPress < DL_HUC_ZERO) THEN
    fConverted := DL_HUC_ZERO;                     // 饱和压异常：结果不可信 / Abnormal saturation pressure
    fSatPress  := DL_HUC_ZERO;
    eErrCode   := E_DL_HumConvErr.eNonFinite;      // 故障级码 / Fault-level code
    RETURN;
END_IF

FC_DL_HumidityUnitConvert := TRUE;                 // 换算有效 / Conversion valid

END_FUNCTION

(* ---- FC_DL_InterpHoldLast.st ---- *)
(*==============================================================================
 * 组件名称 (Component)  : FC_DL_InterpHoldLast
 * 所属子库 (Sublibrary) : DL_MathData
 * 当前版本 (Version)    : 1.0.0
 * 兼容性   (Platform)   : CODESYS 3.5+ / TwinCAT 3 / 汇川 InoProShop / 施耐德 Machine Expert
 *                         仅依赖 IEC 61131-3 标准数学（ABS / MIN / MAX），零厂商私有库
 * 功能描述 (Function)   : 保持型查表（clamp / hold-at-ends 语义）：区间内线性插值，
 *                         **超出末节点保持末节点值，低于首节点保持首节点值，绝不外推**。
 *                         与 FC_DL_InterpTwoPointSlope（可受限外推）形成互补：
 *                         凡是外推会产出无物理意义值（负压力、负流量、超量程阀位）的场合，
 *                         一律用本件，宁可饱和到端点也不产生越界数。
 *                         用途：量程上下限饱和映射、传感器特性表端点延拓、执行器输出限幅映射。
 * 接口     (Interface)  : 输入 afX 升序节点表 [X 单位]、afY 对应值表 [Y 单位]、
 *                         iCount 有效点数 [个]（2..32）、fXin 查询点 [X 单位]；
 *                         输出 fYout 结果（恒在 [afY[1], afY[iCount]] 的包络内） [Y 单位]、
 *                         iSeg 区间下标（越界时为 1 或 iCount-1）[-]、
 *                         bHeld 是否发生端点保持、eErrCode（E_DL_InterpHoldErr）；
 *                         返回值 = bValid 结果可信标志（TRUE = fYout 可信）。
 * 边界     (Boundary)   : ① 属主边界：只做保持型查表，**不做外推**（外推归 TwoPointSlope 件）。
 *                         ② 点数域闸 2..32；越域 → 故障级 eBadCount。
 *                         ③ 非有限双判：查询点 + afX 与 afY **两表**全部元素逐项枚举
 *                         （只查 afX 或只查 afY 都会让插值静默产出非有限值）。
 *                         ④ 段宽近似零 → 比例置 0（取左端值）并置信息级 eDegenerateSeg。
 *                         ⑤ 单调性校验：命中区间两端必须满足 afX[i] <= afX[i+1]，
 *                         违反 → 故障级 eTableNotAsc（不假设强序）。
 *                         ⑥ 结果复检：fYout 必须非有限外，且必须落在两端 afY 的闭包内
 *                         （插值性质保证，越出即说明表或比例异常 → eInternal）。
 *                         ⑦ 零全局耦合（无 GVL / VAR_EXTERNAL / 物理地址）。
 * 分工声明 (Scope)      : 与 `FC_DL_InterpTwoPointSlope` 分工：可外推归那件、保持归本件；
 *                         与 `FC_DL_TableIndexBinarySearch` 分工：定位归那件、取值归本件。
 * 来源标签 (Source Tag) : 原创实现（无外部代码引入）
 * 码表     (Codes)      : 本件不占用全局数字码位；出口为 BOOL + LREAL + INT + BOOL +
 *                         本文件内定义 enum E_DL_InterpHoldErr（全库唯一）。
 * 红线自检 (Redline)    : R1 ✓ 零 GVL/VAR_EXTERNAL ｜ R2 ✓ 零 %I/%Q/%M ｜ R3 ✓ 纯 IEC 61131-3
 *                         R4 ✓ 双表全元素非有限双判 + 段宽判零 + 结果包络复检 ｜ R5 ✓ 声明逐行同行双语注释
 *                         R6 N/A（纯函数无状态机） ｜ R7 N/A（无实例调用）
 * 修订历史 (Revision)   : 2026-11-23  v1.0.0  R77 首版（批次 B3 · 序号 6）
 * 验收向量 (Acceptance) : ① afX=[0,10,20], afY=[0,100,200], iCount=3, fXin=15 →
 *                         fYout=150.0, iSeg=2, bHeld=FALSE, eOk, TRUE；
 *                         ② 同上, fXin=100 → fYout=200.0（保持末值）, iSeg=2, bHeld=TRUE, eOk；
 *                         ③ 同上, fXin=-50 → fYout=0.0（保持首值）, iSeg=1, bHeld=TRUE, eOk；
 *                         ④ 同上, fXin=0 → fYout=0.0, iSeg=1, bHeld=FALSE（恰在首节点，非保持）；
 *                         ⑤ afY[2]=NaN → 返回 FALSE, fYout=0, eNonFinite。
 *==============================================================================*)

(*-----------------------------------------------------------------------------
 * 枚举: E_DL_InterpHoldErr（保持型查表错误码，归属 DL_MathData，与本件同文件，全库唯一属主）
 *----------------------------------------------------------------------------*)
TYPE E_DL_InterpHoldErr :
(
    eOk            := 0,   // 信息级：区间内插值完成 / Info: in-range interpolation done
    eDegenerateSeg := 1,   // 信息级：段宽近似零，取左端值 / Info: degenerate segment, left value used
    eBadCount      := 2,   // 故障级：点数越域 / Fault: point count out of domain
    eNonFinite     := 3,   // 故障级：任一入参或表元素非有限 / Fault: any input or table entry non-finite
    eTableNotAsc   := 4,   // 故障级：表不满足升序约定 / Fault: table violates ascending contract
    eInternal      := 9    // 故障级：结果越出端点包络，内部不一致 / Fault: result outside endpoint envelope
);
END_TYPE

FUNCTION FC_DL_InterpHoldLast : BOOL
VAR_INPUT
    afX    : ARRAY[1..32] OF LREAL;  // 升序节点表 [X 单位] / Ascending node table in X
    afY    : ARRAY[1..32] OF LREAL;  // 对应值表 [Y 单位] / Corresponding value table in Y
    iCount : INT;                    // 有效点数（2..32） [个] / Valid point count, 2..32
    fXin   : LREAL;                  // 查询点 [X 单位] / Query value in X
END_VAR
VAR_OUTPUT
    fYout    : LREAL;  // 结果（恒在端点包络内） [Y 单位] / Result always inside endpoint envelope
    iSeg     : INT;    // 区间下标（越界时为端段） [-] / Segment index, end segment when held
    bHeld    : BOOL;   // 是否发生端点保持 [-] / Whether endpoint hold occurred
    eErrCode : E_DL_InterpHoldErr; // 错误码出口 [-] / Error code outlet
END_VAR
VAR
    _i       : INT;    // 循环下标 [-] / Loop index
    _iSeg    : INT;    // 命中区间下标 [-] / Hit segment index
    _bFound  : BOOL;   // 区间命中标志 [-] / Segment found flag
    _bNonFin : BOOL;   // 非有限标志 [-] / Non-finite flag
    _fDen    : LREAL;  // 段宽（分母） [X 单位] / Segment width denominator
    _fRatio  : LREAL;  // 段内比例 [-] / In-segment ratio
    _fLo     : LREAL;  // 端点包络下界 [Y 单位] / Envelope lower bound
    _fHi     : LREAL;  // 端点包络上界 [Y 单位] / Envelope upper bound
END_VAR
VAR CONSTANT
    DL_IHC_CNT_MIN : INT := 2;        // 点数下限 [个] / Count lower bound
    DL_IHC_CNT_MAX : INT := 32;       // 点数上限（数组容量） [个] / Count upper bound
    DL_IHC_TINY    : LREAL := 1.0E-9; // 段宽近似零阈值 [-] / Degenerate segment threshold
    DL_IHC_ZERO    : LREAL := 0.0;    // 零与比例下限 [-] / Zero and ratio lower bound
    DL_IHC_ONE     : LREAL := 1.0;    // 比例上限 [-] / Ratio upper bound
END_VAR

(* —— 段 0：出口预置安全值 —— *)
FC_DL_InterpHoldLast := FALSE;                     // 返回值预置无效 / Return preset invalid
fYout    := DL_IHC_ZERO;                           // 结果哨兵 0 / Result sentinel
iSeg     := 0;                                     // 下标哨兵 / Index sentinel
bHeld    := FALSE;                                 // 保持标志预置否 / Hold flag preset false
eErrCode := E_DL_InterpHoldErr.eBadCount;          // 预置最严码 / Preset strictest code

(* —— 段 1：点数域闸 —— *)
IF (iCount < DL_IHC_CNT_MIN) OR (iCount > DL_IHC_CNT_MAX) THEN
    RETURN;
END_IF

(* —— 段 2：非有限域闸（查询点 + afX 与 afY 双表逐项枚举） —— *)
_bNonFin := (fXin <> fXin) OR ((fXin - fXin) <> DL_IHC_ZERO);
_i := 1;
WHILE _i <= iCount DO
    IF (afX[_i] <> afX[_i]) OR ((afX[_i] - afX[_i]) <> DL_IHC_ZERO) THEN
        _bNonFin := TRUE;                          // X 表元素非有限 / X entry non-finite
    END_IF
    IF (afY[_i] <> afY[_i]) OR ((afY[_i] - afY[_i]) <> DL_IHC_ZERO) THEN
        _bNonFin := TRUE;                          // Y 表元素非有限 / Y entry non-finite
    END_IF
    _i := _i + 1;
END_WHILE
IF _bNonFin THEN
    eErrCode := E_DL_InterpHoldErr.eNonFinite;
    RETURN;
END_IF

(* —— 段 3：端点保持分支（低于首节点 / 高于末节点，均不外推） —— *)
IF fXin < afX[1] THEN
    fYout    := afY[1];                            // 保持首节点值 / Hold first node value
    iSeg     := 1;
    bHeld    := TRUE;
    eErrCode := E_DL_InterpHoldErr.eOk;
    FC_DL_InterpHoldLast := TRUE;
    RETURN;
END_IF
IF fXin > afX[iCount] THEN
    fYout    := afY[iCount];                       // 保持末节点值 / Hold last node value
    iSeg     := iCount - 1;
    bHeld    := TRUE;
    eErrCode := E_DL_InterpHoldErr.eOk;
    FC_DL_InterpHoldLast := TRUE;
    RETURN;
END_IF

(* —— 段 4：区间定位（升序：afX[i] <= fXin <= afX[i+1]） —— *)
_i      := 1;
_bFound := FALSE;
_iSeg   := 1;
WHILE (_i < iCount) AND (NOT _bFound) DO
    IF (fXin >= afX[_i]) AND (fXin <= afX[_i + 1]) THEN
        _bFound := TRUE;
        _iSeg   := _i;                             // 记录命中区间 / Record hit segment
    ELSE
        _i := _i + 1;
    END_IF
END_WHILE
IF NOT _bFound THEN
    eErrCode := E_DL_InterpHoldErr.eTableNotAsc;   // 未命中：表不满足升序 / Not found: table not ascending
    RETURN;
END_IF

(* —— 段 5：区间升序复检 + 段内比例计算（段宽判零） —— *)
IF afX[_iSeg + 1] < afX[_iSeg] THEN
    eErrCode := E_DL_InterpHoldErr.eTableNotAsc;   // 端点倒序 / Endpoints reversed
    RETURN;
END_IF
_fDen := afX[_iSeg + 1] - afX[_iSeg];              // 段宽 / Segment width
IF ABS(_fDen) < DL_IHC_TINY THEN
    _fRatio  := DL_IHC_ZERO;                       // 退化段取左端 / Degenerate: use left node
    eErrCode := E_DL_InterpHoldErr.eDegenerateSeg; // 信息级码 / Info code
ELSE
    _fRatio  := (fXin - afX[_iSeg]) / _fDen;       // 标准比例 / Standard ratio
    eErrCode := E_DL_InterpHoldErr.eOk;            // 信息级成功 / Info success
END_IF
_fRatio := MIN(MAX(_fRatio, DL_IHC_ZERO), DL_IHC_ONE);   // 显式约束 0..1 / Constrain 0..1

(* —— 段 6：线性插值取值 —— *)
fYout := afY[_iSeg] + (afY[_iSeg + 1] - afY[_iSeg]) * _fRatio;
iSeg  := _iSeg;
bHeld := FALSE;                                    // 区间内不属保持 / In-range, not a hold

(* —— 段 7：结果复检（非有限 + 端点包络） —— *)
IF (fYout <> fYout) OR ((fYout - fYout) <> DL_IHC_ZERO) THEN
    fYout    := DL_IHC_ZERO;
    iSeg     := 0;
    eErrCode := E_DL_InterpHoldErr.eNonFinite;
    RETURN;
END_IF
_fLo := MIN(afY[_iSeg], afY[_iSeg + 1]);           // 包络下界 / Envelope lower bound
_fHi := MAX(afY[_iSeg], afY[_iSeg + 1]);           // 包络上界 / Envelope upper bound
IF (fYout < _fLo) OR (fYout > _fHi) THEN
    fYout    := DL_IHC_ZERO;                       // 越出包络：内部不一致 / Outside envelope: internal fault
    iSeg     := 0;
    eErrCode := E_DL_InterpHoldErr.eInternal;
    RETURN;
END_IF

FC_DL_InterpHoldLast := TRUE;                      // 结果有效 / Result valid

END_FUNCTION

(* ---- FC_DL_InterpLogLinear.st ---- *)
(*==============================================================================
 * 组件名称 (Component)  : FC_DL_InterpLogLinear
 * 所属子库 (Sublibrary) : DL_MathData
 * 当前版本 (Version)    : 1.0.0
 * 兼容性   (Platform)   : CODESYS 3.5+ / TwinCAT 3 / 汇川 InoProShop / 施耐德 Machine Expert
 *                         仅依赖 IEC 61131-3 标准数学（LN / ABS），零厂商私有库
 * 功能描述 (Function)   : 对数-线性插值（X 取对数、Y 线性）：跨数量级工艺曲线插值。
 *                           y = y1 + (y2 - y1) × (LN(x) - LN(x1)) / (LN(x2) - LN(x1))
 *                         典型用途：流量-压差（孔板特性）、风机风量-静压、传感器对数刻度。
 *                         **适用域**：x1 > 0 且 x2 > 0 且 xin > 0（对数定义域），
 *                         任一为 0 或负 → 故障级 eOutOfLogDomain，**不静默取绝对值**。
 *                         xin 允许落在 [x1, x2] 之外的近邻区（线性于对数域外推），
 *                         但外推幅度受 fExtrapRatio 上限（默认 1.0，即最多外推一个
 *                         对数区间的宽度）钳制；超限钳位并置信息级 eExtrapClamped。
 * 接口     (Interface)  : 输入 fX1/fY1 左节点、fX2/fY2 右节点、fXin 查询点、
 *                         fExtrapRatio 允许的最大外推比例 [倍数，默认 1.0]；
 *                         输出 fYout 插值结果 [Y 单位]、fSel 实际使用的对数域位置比 [0..1+外推]、
 *                         bExtrapolated 是否发生外推、eErrCode（E_DL_InterpLogErr）；
 *                         返回值 = bValid 插值可信标志（TRUE = fYout 可信）。
 * 边界     (Boundary)   : ① 属主边界：只做两点对数-线性插值，不做多点表遍历（表遍历归查表族）。
 *                         ② 全浮点入参（5 个）非有限双判，逐一枚举，漏一个即静默失效。
 *                         ③ 对数域闸：x1 <= 0 或 x2 <= 0 或 xin <= 0 → 故障级 eOutOfLogDomain。
 *                         ④ 对数区间宽度判零：|LN(x2)-LN(x1)| < 1E-12 → 故障级 eDegenerateSeg
 *                         （两节点 X 相同，插值无定义），避免除零。
 *                         ⑤ 外推上限：fExtrapRatio <= 0 视为非法参数 → 故障级 eBadParam。
 *                         ⑥ 零全局耦合（无 GVL / VAR_EXTERNAL / 物理地址）。
 * 分工声明 (Scope)      : 与 `FC_DL_InterpTwoPointSlope` 分工：线性斜率外推归那件、
 *                         对数域插值归本件；与 `FC_DL_InterpHoldLast` 分工：保持型归那件。
 * 来源标签 (Source Tag) : 原创实现（无外部代码引入）
 * 码表     (Codes)      : 本件不占用全局数字码位；出口为 BOOL + 2×LREAL + BOOL +
 *                         本文件内定义 enum E_DL_InterpLogErr（全库唯一）。
 * 红线自检 (Redline)    : R1 ✓ 零 GVL/VAR_EXTERNAL ｜ R2 ✓ 零 %I/%Q/%M ｜ R3 ✓ 纯 IEC 61131-3
 *                         R4 ✓ 全入参非有限双判 + 对数域闸 + 对数区间判零 + 外推钳位 ｜ R5 ✓ 声明逐行同行双语注释
 *                         R6 N/A（纯函数无状态机） ｜ R7 N/A（无实例调用）
 * 修订历史 (Revision)   : 2026-11-23  v1.0.0  R77 首版（批次 B3 · 序号 3）
 * 验收向量 (Acceptance) : ① fX1=1, fY1=0, fX2=10, fY2=100, fXin=3.16227766（=√10）, fExtrapRatio=1.0 →
 *                         LN 位置比 = LN(3.16227766)/LN(10) = 0.5 → fYout = 50.0（容差 1E-6）；
 *                         ② 同上, fXin=1.0 → 位置比 0 → fYout = 0.0, bExtrapolated=FALSE；
 *                         ③ fX1=0 → 返回 FALSE, fYout=0, eOutOfLogDomain；
 *                         ④ fX1=5, fX2=5（区间退化）→ 返回 FALSE, eDegenerateSeg；
 *                         ⑤ fExtrapRatio=0.0 → 返回 FALSE, eBadParam。
 *==============================================================================*)

(*-----------------------------------------------------------------------------
 * 枚举: E_DL_InterpLogErr（对数-线性插值错误码，归属 DL_MathData，与本件同文件，全库唯一属主）
 *----------------------------------------------------------------------------*)
TYPE E_DL_InterpLogErr :
(
    eOk             := 0,   // 信息级：插值完成，无外推 / Info: interpolated, no extrapolation
    eExtrapolated   := 1,   // 信息级：发生受限外推 / Info: bounded extrapolation performed
    eExtrapClamped  := 2,   // 信息级：外推超限已钳位 / Info: extrapolation clamped to limit
    eOutOfLogDomain := 3,   // 故障级：X 非正，超出对数定义域 / Fault: non-positive X, outside log domain
    eDegenerateSeg  := 4,   // 故障级：对数区间宽度为零 / Fault: zero log interval width
    eBadParam       := 5,   // 故障级：外推比例参数非法 / Fault: illegal extrapolation ratio parameter
    eNonFinite      := 6    // 故障级：入参非有限 / Fault: non-finite input
);
END_TYPE

FUNCTION FC_DL_InterpLogLinear : BOOL
VAR_INPUT
    fX1         : LREAL;  // 左节点 X（必须 > 0） [X 单位] / Left node X, must be positive
    fY1         : LREAL;  // 左节点 Y [Y 单位] / Left node Y
    fX2         : LREAL;  // 右节点 X（必须 > 0） [X 单位] / Right node X, must be positive
    fY2         : LREAL;  // 右节点 Y [Y 单位] / Right node Y
    fXin        : LREAL;  // 查询点（必须 > 0） [X 单位] / Query X, must be positive
    fExtrapRatio: LREAL;  // 允许的最大外推比例（对数区间宽度的倍数） [倍数] / Allowed extrapolation ratio
END_VAR
VAR_OUTPUT
    fYout         : LREAL;  // 插值结果 [Y 单位] / Interpolated result
    fSel          : LREAL;  // 对数域位置比（0 = 左节点，1 = 右节点） [-] / Position ratio in log domain
    bExtrapolated : BOOL;   // 是否发生外推 [-] / Whether extrapolation occurred
    eErrCode      : E_DL_InterpLogErr; // 错误码出口 [-] / Error code outlet
END_VAR
VAR
    _bNonFin : BOOL;   // 入参非有限标志 [-] / Non-finite input flag
    _fL1     : LREAL;  // 左节点自然对数 [-] / Natural log of left node
    _fL2     : LREAL;  // 右节点自然对数 [-] / Natural log of right node
    _fLin    : LREAL;  // 查询点自然对数 [-] / Natural log of query
    _fDen    : LREAL;  // 对数区间宽度（分母） [-] / Log interval width denominator
    _fPos    : LREAL;  // 未钳位位置比 [-] / Raw position ratio
    _fLo     : LREAL;  // 位置比下界（负外推上限） [-] / Position lower bound
    _fHi     : LREAL;  // 位置比上界（正外推上限） [-] / Position upper bound
END_VAR
VAR CONSTANT
    DL_ILC_ZERO : LREAL := 0.0;    // 零与位置比左端 [-] / Zero and ratio origin
    DL_ILC_ONE  : LREAL := 1.0;    // 位置比右端 [-] / Ratio at right node
    DL_ILC_TINY : LREAL := 1.0E-12; // 对数区间宽度近似零阈值 [-] / Degenerate log width threshold
END_VAR

(* —— 段 0：出口预置安全值 —— *)
FC_DL_InterpLogLinear := FALSE;                    // 返回值预置无效 / Return preset invalid
fYout         := DL_ILC_ZERO;                      // 结果哨兵 0 / Result sentinel
fSel          := DL_ILC_ZERO;                      // 位置比哨兵 0 / Ratio sentinel
bExtrapolated := FALSE;                            // 外推标志预置否 / Extrapolation preset false
eErrCode      := E_DL_InterpLogErr.eBadParam;      // 预置最严码 / Preset strictest code

(* —— 段 1：非有限域闸（5 个浮点入参逐一枚举） —— *)
_bNonFin := (fX1 <> fX1) OR ((fX1 - fX1) <> DL_ILC_ZERO);            // X1 非有限 / X1 non-finite
_bNonFin := _bNonFin OR (fY1 <> fY1) OR ((fY1 - fY1) <> DL_ILC_ZERO); // Y1 非有限 / Y1 non-finite
_bNonFin := _bNonFin OR (fX2 <> fX2) OR ((fX2 - fX2) <> DL_ILC_ZERO); // X2 非有限 / X2 non-finite
_bNonFin := _bNonFin OR (fY2 <> fY2) OR ((fY2 - fY2) <> DL_ILC_ZERO); // Y2 非有限 / Y2 non-finite
_bNonFin := _bNonFin OR (fXin <> fXin) OR ((fXin - fXin) <> DL_ILC_ZERO);   // X 查询非有限 / Query non-finite
_bNonFin := _bNonFin OR (fExtrapRatio <> fExtrapRatio) OR ((fExtrapRatio - fExtrapRatio) <> DL_ILC_ZERO); // 外推比非有限
IF _bNonFin THEN
    eErrCode := E_DL_InterpLogErr.eNonFinite;      // 故障级码 / Fault-level code
    RETURN;
END_IF

(* —— 段 2：对数域闸（三个 X 均须严格为正） —— *)
IF (fX1 <= DL_ILC_ZERO) OR (fX2 <= DL_ILC_ZERO) OR (fXin <= DL_ILC_ZERO) THEN
    eErrCode := E_DL_InterpLogErr.eOutOfLogDomain; // 故障级：超出对数定义域 / Fault: outside log domain
    RETURN;
END_IF

(* —— 段 3：外推比例参数域闸（必须 > 0，否则外推窗无意义） —— *)
IF fExtrapRatio <= DL_ILC_ZERO THEN
    eErrCode := E_DL_InterpLogErr.eBadParam;       // 故障级：参数非法 / Fault: illegal parameter
    RETURN;
END_IF

(* —— 段 4：对数区间宽度计算与判零（防除零） —— *)
_fL1  := LN(fX1);                                  // 左节点对数 / Log of left node
_fL2  := LN(fX2);                                  // 右节点对数 / Log of right node
_fLin := LN(fXin);                                 // 查询点对数 / Log of query
_fDen := _fL2 - _fL1;                              // 对数区间宽度 / Log interval width
IF ABS(_fDen) < DL_ILC_TINY THEN
    eErrCode := E_DL_InterpLogErr.eDegenerateSeg;  // 故障级：区间退化 / Fault: degenerate interval
    RETURN;                                        // 早退，杜绝除零 / Early exit, avoids division by zero
END_IF

(* —— 段 5：位置比计算与受限外推钳位 —— *)
_fPos := (_fLin - _fL1) / _fDen;                   // 对数域位置比 / Position ratio in log domain
_fLo  := DL_ILC_ZERO - fExtrapRatio;               // 负外推上限 / Lower extrapolation bound
_fHi  := DL_ILC_ONE + fExtrapRatio;                // 正外推上限 / Upper extrapolation bound

IF _fPos < DL_ILC_ZERO THEN
    bExtrapolated := TRUE;                         // 负向外推 / Negative extrapolation
    IF _fPos < _fLo THEN
        _fPos    := _fLo;                          // 外推超限钳位 / Clamp extrapolation
        eErrCode := E_DL_InterpLogErr.eExtrapClamped;
    ELSE
        eErrCode := E_DL_InterpLogErr.eExtrapolated;
    END_IF
ELSIF _fPos > DL_ILC_ONE THEN
    bExtrapolated := TRUE;                         // 正向外推 / Positive extrapolation
    IF _fPos > _fHi THEN
        _fPos    := _fHi;                          // 外推超限钳位 / Clamp extrapolation
        eErrCode := E_DL_InterpLogErr.eExtrapClamped;
    ELSE
        eErrCode := E_DL_InterpLogErr.eExtrapolated;
    END_IF
ELSE
    bExtrapolated := FALSE;                        // 区间内正常插值 / Normal in-range interpolation
    eErrCode      := E_DL_InterpLogErr.eOk;
END_IF

(* —— 段 6：插值取值 —— *)
fYout       := fY1 + (fY2 - fY1) * _fPos;          // y = y1 + (y2-y1)*位置比 / Linear in Y over log position
fSel        := _fPos;                              // 导出位置比 / Export position ratio

(* —— 段 7：结果非有限复检兜底 —— *)
IF (fYout <> fYout) OR ((fYout - fYout) <> DL_ILC_ZERO) THEN
    fYout    := DL_ILC_ZERO;                       // 复检异常回哨兵 / Recheck failed: sentinel
    fSel     := DL_ILC_ZERO;
    eErrCode := E_DL_InterpLogErr.eNonFinite;      // 故障级码 / Fault-level code
    RETURN;
END_IF

FC_DL_InterpLogLinear := TRUE;                     // 插值有效 / Interpolation valid

END_FUNCTION
